(* IEC 61131-3 sources: daoli-st-library/DL_Motion (part 13) *)

(* ---- FB_DL_FilmWebCenter.st ---- *)
(*
    FB_DL_FilmWebCenter —— 膜卷纠偏（EPC）
    ------------------------------------------------------------------
    分类      : DL_Motion / Guide
    前缀      : FB_DL_
    版本      : 1.0.0
    溯源      : 纠偏为公开卷材处理工程结构（EPC / CPC：边缘或中心偏差 → 纠偏辊位置给定）；
                死区保持、断料保持、限速率、双侧行程钳位、错误分级与码位 100% 自有；
                与排线往复件、背隙修正件的职责严格分离（一个管横向对中、一个管往复排布、
                一个管传动链间隙）；clean-room 重写，未复制任何闭源厂商源码
    平台      : 纯 IEC 61131-3，CODESYS V3.5+ / TwinCAT 3 / InoProShop 通用
    作者      : 道莅代码库 · PLC编程专家（R19）
    ------------------------------------------------------------------
    功能说明  : 把边缘/中心偏差换算成纠偏辊位置给定。核心防御三条：
                ① 死区内保持——偏差在死区内给定不动，防辊子随噪声来回磨（不是把给定设成 0）；
                ② 限速率——纠偏动作过快会造成膜起皱甚至跑偏振荡；
                ③ 断料保持——膜断了还继续纠偏，辊子会一路顶到机械极限，复产后第一次穿膜
                   直接撞限位，故断料时给定保持末值、绝不追 0。
                其余防御：④ 行程域矛盾、增益或速率越域即故障级 02E4 并冻结在中心位
                   （增益过大是纠偏振荡的头号原因，硬限比「相信现场」更安全）；
                ⑤ 偏差非有限即故障级 02E5 并保持末次给定；
                ⑥ 给定双侧行程钳位，超限置 bLimited；⑦ 斜率限制首拍 fStep 由引脚换算，
                   不做除法；⑧ 状态机 CASE 含 ELSE 兜底，非法状态回 eIdle 并保持给定。
                职责边界：纠偏执行器的伺服闭环归驱动层，本件只出位置给定。
    错误码    : 16#0004_01D1 断料保持中 / 偏差在死区内给定保持——信息级，正常防御
                16#0004_01D2 预留禁用（信息级，不得挪用）
                16#0004_02E4 增益/速率/行程/采样参数非法——故障级，纠偏冻结在中心位
                16#0004_02E5 偏差输入非有限——故障级，给定保持末次有效
                16#0004_02E6 状态机落 ELSE 兜底（非法状态）——故障级，回 eIdle 并保持给定
    码位总账  : 16#0004_01D1 用 / 16#0004_01D2 预留 ｜ 16#0004_02E4 用 / 16#0004_02E5 用 / 16#0004_02E6 用
    状态机    : E_DL_WebState（eIdle / eManual / eAuto / eWebLost / eFault）五态，CASE 含 ELSE 兜底，
                ELSE 回 eIdle 并置故障级 02E6；失能不归零，只保持末值。
    采样约定  : fbTrigReset 在本体首部无条件刷新；速率步长由 tSampleTime 引脚换算；
                bInDeadband / bLimited / bWebLost 均为当拍组合量，不锁存。
    修订记录  : 2026-11-16 v1.0.0 首次入库（R19）
*)

(*
    枚举 : E_DL_WebState —— 纠偏工作状态（本文件为全库唯一属主）
*)
TYPE E_DL_WebState :
(
    eIdle    := 0,                            // 空闲：未使能，给定保持 / idle, disabled, the setpoint is held
    eManual  := 1,                            // 手动：走手动偏置给定 / manual, the setpoint follows the manual offset
    eAuto    := 2,                            // 自动：按偏差纠偏 / automatic, correcting by the measured deviation
    eWebLost := 3,                            // 断料：给定保持末值 / web lost, the setpoint holds its last value
    eFault   := 4                             // 故障：冻结在中心位 / fault, frozen at the centre
);
END_TYPE

FUNCTION_BLOCK FB_DL_FilmWebCenter
VAR_INPUT
    bEnable         : BOOL;                   // 使能，FALSE 输出保持末值（不归零）/ enable, FALSE holds the last setpoint without zeroing it
    bReset          : BOOL;                   // 复位，上升沿回中位并清状态 / reset, rising edge returns to the centre and clears the state
    bAuto           : BOOL := FALSE;          // TRUE = 自动纠偏，FALSE = 手动（走 fManualOffset）/ TRUE automatic, FALSE manual via the manual offset
    fDeviation      : REAL := 0.0;            // 边缘/中心偏差（正 = 偏向驱动侧）[mm] / edge or centre deviation, positive towards the drive side [mm]
    fGain           : REAL := 1.0;            // 偏差到位置给定增益 [mm/mm]，范围 0.1~20.0 / deviation to position gain [mm/mm], range 0.1~20.0
    fManualOffset   : REAL := 0.0;            // 手动偏置 [mm]，范围 fTravelMin~fTravelMax / manual offset [mm], range fTravelMin~fTravelMax
    fDeadband       : REAL := 0.3;            // 死区半宽 [mm]，范围 0.0~10.0 / deadband half width [mm], range 0.0~10.0
    fRateMax        : REAL := 5.0;            // 给定最大变化率 [mm/s]，范围 0.01~100.0 / maximum setpoint rate [mm/s], range 0.01~100.0
    fTravelMin      : REAL := -50.0;          // 行程下限 [mm] / travel lower bound [mm]
    fTravelMax      : REAL := 50.0;           // 行程上限 [mm]，必须 > fTravelMin / travel upper bound [mm], must be > fTravelMin
    bWebPresent     : BOOL := TRUE;           // 膜在位信号，FALSE = 断料 / web present signal, FALSE means the web is lost
    tSampleTime     : TIME := T#20MS;         // 采样周期 [ms]，范围 1~1000 / sample time [ms], range 1~1000
END_VAR
VAR_OUTPUT
    fPositionSp     : REAL;                   // 纠偏辊位置给定 [mm] / guide roller position setpoint [mm]
    bInDeadband     : BOOL;                   // 偏差在死区内（给定保持）/ the deviation is inside the deadband, the setpoint holds
    bLimited        : BOOL;                   // 受行程或速率限制 / limited by the travel or the rate
    bWebLost        : BOOL;                   // 断料保持中 / holding because the web is lost
    eErr            : UDINT;                  // 错误码，0=正常 / error id, 0=ok
    bError          : BOOL;                   // 故障标志，eErr 为故障级时 TRUE / error flag, TRUE on fault-level eErr
    bValid          : BOOL;                   // 给定是否可用 / setpoint valid flag
END_VAR
VAR
    fbTrigReset     : R_TRIG;                 // 复位上升沿实例，本体首部无条件刷新 / reset edge instance, refreshed unconditionally
    eState          : E_DL_WebState := eIdle; // 状态机当前态 / current state machine state
    fLastSp         : REAL;                   // 上一拍给定（斜率基准）[mm] / previous setpoint used by the ramp [mm]
    fTarget         : REAL;                   // 钳位与限速率前的目标给定 [mm] / target setpoint before clamping and ramping [mm]
    fStep           : REAL;                   // 本拍允许的最大变化量 [mm] / maximum allowed change in this cycle [mm]
    fDtSec          : REAL;                   // 采样周期秒值 [s] / sample time in seconds [s]
    fGainEff        : REAL;                   // 钳位后的增益 [mm/mm] / clamped gain [mm/mm]
    fDeadEff        : REAL;                   // 钳位后的死区半宽 [mm] / clamped deadband half width [mm]
    fManualEff      : REAL;                   // 钳位后的手动偏置 [mm] / clamped manual offset [mm]
    nDtMs           : DINT;                   // 采样周期毫秒整数 [ms] / sample time in integer milliseconds [ms]
    bInit           : BOOL := FALSE;          // 首扫标志，初值 FALSE，判据 NOT bInit / first-scan flag, initial FALSE, tested with NOT
END_VAR
VAR CONSTANT
    DL_EPC_GAIN_MIN  : REAL := 0.1;           // 增益下限 [mm/mm] / gain lower bound [mm/mm]
    DL_EPC_GAIN_MAX  : REAL := 20.0;          // 增益上限 [mm/mm] / gain upper bound [mm/mm]
    DL_EPC_RATE_MIN  : REAL := 0.01;          // 速率下限 [mm/s] / rate lower bound [mm/s]
    DL_EPC_RATE_MAX  : REAL := 100.0;         // 速率上限 [mm/s] / rate upper bound [mm/s]
    DL_EPC_DB_MAX    : REAL := 10.0;          // 死区半宽上限 [mm] / deadband half width upper bound [mm]
    DL_EPC_DT_MAX    : TIME := T#1S;          // 采样周期上限 [ms] / sample time upper bound [ms]
    DL_EPC_DT_MIN    : TIME := T#1MS;         // 采样周期下限 [ms] / sample time lower bound [ms]
    DL_FLOAT_EPS     : REAL := 1.0E-6;        // 浮点判等容差 [无量纲] / float equality tolerance [dimensionless]
    DL_EPC_MS_PER_S  : REAL := 1000.0;        // 毫秒到秒换算因子 [ms/s] / milliseconds per second [ms/s]
    DL_EPC_INF_GUARD : REAL := 1.0E38;        // 非有限幅值判定阈值 [无量纲] / non-finite magnitude guard [dimensionless]
    DL_EPC_ZERO      : REAL := 0.0;           // 零值常量，避免裸字面量 [mm] / zero constant, avoids a bare literal [mm]
END_VAR

// 段 1｜边沿实例无条件周期刷新（红线：严禁放入条件分支）/ segment 1, unconditional edge refresh
fbTrigReset(CLK := bReset);

// 段 2｜输出与错误状态预置（fPositionSp 为保持量，故障与断料时均保持）/ segment 2, preset outputs, the setpoint is held
eErr := 0;                                    // 预置无错误 / preset no error
bError := FALSE;                              // 预置无故障 / preset no fault
bInDeadband := FALSE;                         // 预置非死区 / preset outside the deadband
bLimited := FALSE;                            // 预置未受限 / preset not limited
bWebLost := NOT bWebPresent;                  // 断料标志由在位信号导出 / the web lost flag derives from the present signal

// 段 3｜首扫初始化（唯一合法范式：初值 FALSE，判据 NOT bInit）/ segment 3, first-scan initialisation
IF NOT bInit THEN
    fLastSp := DL_EPC_ZERO;                   // 首扫给定基准取中心位 / the setpoint reference starts at the centre
    bInit := TRUE;                            // 首扫只做一次 / first scan runs once only
END_IF

// 段 4｜参数闸：行程域、增益、速率、采样周期（任一非法即冻结在中心位）/ segment 4, parameter gate
IF (fTravelMax <= fTravelMin)
   OR (fGain < DL_EPC_GAIN_MIN) OR (fGain > DL_EPC_GAIN_MAX)
   OR (fRateMax < DL_EPC_RATE_MIN) OR (fRateMax > DL_EPC_RATE_MAX)
   OR (tSampleTime < DL_EPC_DT_MIN) OR (tSampleTime > DL_EPC_DT_MAX) THEN
    eErr := 16#0004_02E4;                     // 参数非法故障码 / illegal parameter fault id
    bError := TRUE;                           // 置故障标志 / raise the error flag
    eState := eFault;                         // 落故障态 / enter the fault state
    fPositionSp := DL_EPC_ZERO;               // 冻结在中心位（唯一安全的固定点）/ freeze at the centre, the only safe fixed point
    bValid := FALSE;                          // 给定不可用 / the setpoint is not usable
    RETURN;                                   // 故障级提前返回 / early return on fault
END_IF

// 段 5｜偏差非有限闸：给定保持末次有效（绝不追 0）/ segment 5, non-finite gate holds the setpoint
IF (fDeviation <> fDeviation) OR (fDeviation > DL_EPC_INF_GUARD) OR (fDeviation < -DL_EPC_INF_GUARD) THEN
    eErr := 16#0004_02E5;                     // 偏差非有限故障码 / non-finite deviation fault id
    bError := TRUE;                           // 置故障标志 / raise the error flag
    eState := eFault;                         // 落故障态 / enter the fault state
    fPositionSp := fLastSp;                   // 保持末次给定 / hold the last setpoint
    bValid := FALSE;                          // 给定不可用 / the setpoint is not usable
    RETURN;                                   // 故障级提前返回 / early return on fault
END_IF

// 段 6｜域钳位与速率步长（无历史依赖，不做除法）/ segment 6, domain clamp and rate step
fGainEff := fGain;                            // 增益已由段 4 保证在域内 / the gain is already in range by segment 4
fDeadEff := MIN(MAX(fDeadband, DL_EPC_ZERO), DL_EPC_DB_MAX); // 死区半宽收敛到 0.0~10.0 mm / converge the deadband into 0.0~10.0 mm
fManualEff := MIN(MAX(fManualOffset, fTravelMin), fTravelMax); // 手动偏置收敛到行程域 / converge the manual offset into the travel range
nDtMs := TIME_TO_DINT(tSampleTime);           // 采样周期整数毫秒 [ms] / sample time in integer milliseconds [ms]
fDtSec := DINT_TO_REAL(nDtMs) / DL_EPC_MS_PER_S; // 换算为秒，除子为常量 [s] / convert to seconds, the divisor is a constant [s]
fStep := fRateMax * fDtSec;                   // 本拍允许的最大变化量 [mm] / maximum allowed change in this cycle [mm]

// 段 7｜复位沿：回中位并清状态 / segment 7, reset returns to the centre
IF fbTrigReset.Q THEN
    fLastSp := DL_EPC_ZERO;                   // 给定基准回中心位 / the setpoint reference returns to the centre
    fPositionSp := DL_EPC_ZERO;               // 给定回中位 / the setpoint returns to the centre
    IF eState = eFault THEN
        eState := eIdle;                      // 故障态允许由复位退出 / a reset leaves the fault state
    END_IF
END_IF

// 段 8｜状态选择（断料优先级最高，其次使能与手自动）/ segment 8, state selection
IF NOT bWebPresent THEN
    eState := eWebLost;                       // 断料优先，给定保持 / web loss has the highest priority, the setpoint holds
    bWebLost := TRUE;                         // 发布断料标志 / publish the web lost flag
ELSE
    bWebLost := FALSE;                        // 在位则清断料标志 / clear the flag when the web is present
    IF eState = eWebLost THEN
        eState := eIdle;                      // 断料解除回空闲，由使能重新决定手自动 / leaving the web lost state returns to idle
    END_IF
END_IF
IF (eState <> eWebLost) AND (eState <> eFault) THEN
    IF NOT bEnable THEN
        eState := eIdle;                      // 失能回空闲（保持不归零）/ disabled returns to idle without zeroing the setpoint
    ELSIF bAuto THEN
        eState := eAuto;                      // 自动纠偏 / automatic correction
    ELSE
        eState := eManual;                    // 手动偏置 / manual offset
    END_IF
END_IF

// 段 9｜目标给定（含死区保持与断料保持）/ segment 9, target setpoint with deadband and web loss holding
CASE eState OF
    eIdle:
        fTarget := fLastSp;                   // 空闲保持末值，不归零 / idle holds the last value without zeroing it

    eManual:
        fTarget := fManualEff;                // 手动走偏置给定 / manual follows the offset

    eAuto:
        IF ABS(fDeviation) <= fDeadEff THEN
            fTarget := fLastSp;               // 死区内保持，绝不设成 0 / hold inside the deadband, never set it to zero
            bInDeadband := TRUE;              // 发布死区标志 / publish the deadband flag
            eErr := 16#0004_01D1;             // 信息级：偏差在死区内给定保持 / info level, the setpoint holds inside the deadband
        ELSE
            fTarget := fLastSp + fGainEff * fDeviation; // 增量式纠偏：在上一拍给定上叠加 / incremental correction on top of the previous setpoint
        END_IF

    eWebLost:
        fTarget := fLastSp;                   // 断料保持末值 / web lost holds the last value
        eErr := 16#0004_01D1;                 // 信息级：断料保持中 / info level, holding because the web is lost

    eFault:
        fTarget := fLastSp;                   // 故障态保持末值 / the fault state holds the last value

ELSE
    eErr := 16#0004_02E6;                     // 故障级：非法状态兜底 / fault level, illegal state fallback
    bError := TRUE;                           // 置故障标志 / raise the error flag
    eState := eIdle;                          // 回空闲态 / fall back to idle
    fTarget := fLastSp;                       // 保持末值，不产生跳变 / hold the last value, no jump
END_CASE

// 段 10｜行程双侧钳位（只做单侧是常见缺陷）/ segment 10, two-sided travel clamp
IF fTarget > fTravelMax THEN
    fTarget := fTravelMax;                    // 上限钳位 / clamp at the upper bound
    bLimited := TRUE;                         // 标记行程受限 / flag the travel limit
ELSIF fTarget < fTravelMin THEN
    fTarget := fTravelMin;                    // 下限钳位 / clamp at the lower bound
    bLimited := TRUE;                         // 标记行程受限 / flag the travel limit
END_IF

// 段 11｜限速率（每拍最多变化 fStep，防膜起皱与跑偏振荡）/ segment 11, rate limiting
IF fStep > DL_EPC_ZERO THEN
    IF fTarget > (fLastSp + fStep) THEN
        fTarget := fLastSp + fStep;           // 正向每拍限幅 / limit the positive step per cycle
        bLimited := TRUE;                     // 标记速率受限 / flag the rate limit
    ELSIF fTarget < (fLastSp - fStep) THEN
        fTarget := fLastSp - fStep;           // 负向每拍限幅 / limit the negative step per cycle
        bLimited := TRUE;                     // 标记速率受限 / flag the rate limit
    END_IF
END_IF

// 段 12｜发布给定 / segment 12, publish the setpoint
fPositionSp := fTarget;                       // 输出纠偏辊位置给定 [mm] / publish the guide roller setpoint [mm]
fLastSp := fTarget;                           // 记录为下一拍斜率基准 / remember it as the next ramp reference
IF NOT bError THEN
    bValid := TRUE;                           // 无故障则给定可用 / usable when no fault is present
END_IF
END_FUNCTION_BLOCK

(* ---- FB_DL_FlyingCutSync.st ---- *)
(*
  FB_DL_FlyingCutSync  —  飞剪同步切（相位取模 / 切窗判据 / 电子齿轮追赶 / 单拍下刀）/ Flying-cut synchronisation
  分类 Category : DL_Motion
  码位 Code     : 16#04_0_A3
  版本 Version  : 1.0.1
  来源 Source   : t1-6-plcopen — IEC 61131-3 标准语义的道莅防御性实现
  溯源 Origin   : PLCopen 飞剪/电子齿轮公开语义借鉴，clean-room 实现，仅借相位取模与切窗概念，未复制源码行
  功能 Function : 1) 主轴位置对 fCutLengthMm 取模（FLOOR 口径，负向同样收敛）得切长相位 fPhaseMm；
                  2) 相位落在 [fSyncWindowStartMm, fSyncWindowEndMm] 内置 bInSyncWindow，窗口内方允许下刀；
                  3) 同步误差 fSyncErrorMm = 刀轴位置 − 相位 × fCutOverlapRatio，进 fSyncTolMm 才发下刀脉冲；
                  4) 下刀脉冲 bCutCmd 为**单拍脉冲**（脉冲语义：置位 1 个 PLC 周期），由内部 _bCutPulse 置位、
                     段 8 统一出口映射，次拍段 1 清零，绝不在 CASE 内二次写输出（N2 / R187①）；
                  5) 切完按 tCutDwell 保压（刀在料内停留），保压结束进回程相，等相位越过窗尾再回等待相；
                  6) 每圈只允许一刀：以圈索引 fTurnsInt 与 _nCutTurnIdx 比较做单圈互锁（防同圈重刀）。
  边界 Boundary : ① fCutLengthMm <= 0 判组态错（取模除零前置，R45）；窗口起止倒置或宽 <= 0 判组态错且不运行；
                      fSyncTolMm <= 0 / fCutOverlapRatio <= 0 同判组态错，码 00A3，状态进 eFault；
                  ② 未同步时**禁止** bCutCmd：互锁写在件内（窗口 + 容差 + 单圈 + 主轴正向四条件同时成立），
                     不外抛给上层组合逻辑（防上层漏联锁切刀撞料）；
                  ③ nCutCount 到 uCountPreset 后 bPresetReached 置位；计数在 UDINT 上限前饱和**不回绕**，
                     预置比较用「增量前预判」而非事后比较（不给 TRUNC(x)+1 型写法，R28-3）；
                  ④ 切窗内主轴反转立即判废并置 01A3（反转期刀轴与料带速度矢量相反，下刀即撕料）；
                  ⑤ uCountPreset = 0 视为「不启用预置」：bPresetReached 恒 FALSE，置信息级 07A3；
                  ⑥ 解除路径自证：_bFault 清除 = rtReset.Q（引脚可满足）；01A3 另可由「主轴恢复正向
                     且相位出新窗」按码专清（两路径互不掩盖，R188）。
  依赖 Depends  : I_DL_MotionAxis / E_DL_AxisState（DL_Motion 既有契约件，零修改，只注入不实例化）；
                  仅 Standard.library（TON / R_TRIG / ABS / MIN / MAX）
  同拍双窗配比  : tCutDwell（刀内停留）与 tonGuard 自复位心跳窗不同源；配比约束
                  tCutDwell <= DL_GUARD_WINDOW / 2，保证保压段内至少一次心跳判活（R100）

  码表 Error codes（本件格 04_0_A3，子码步进 +0x10）:
    16#0004_00A3 故障级：组态非法（切长 <= 0 / 窗口倒置或宽 <= 0 / 容差 <= 0 / 重叠比 <= 0）
    16#0004_01A3 故障级：切窗内主轴反转，本次切割判废
    16#0004_03A3 故障级：状态机落 ELSE 兜底（非法相位 ID）
    16#0004_04A3 信息级：下刀脉冲已发出（bCutCmd 单拍同源，不置 bError）
    16#0004_05A3 信息级：切割计数达预置（bPresetReached 同拍置位，不置 bError）
    16#0004_06A3 信息级：切窗内同步超差，本次跳过不下刀（互锁生效，不置 bError）
    16#0004_07A3 信息级：预置计数未组态（uCountPreset = 0，预置出口恒 FALSE）

  修订历史 Revision :
    2026-11-18  v1.0.0  R37 首版
*)

TYPE E_DL_FlyingCutState :
(
    eIdle       := 0,   // 空闲：未使能，不出切窗判据 / Idle, no window evaluation while disabled
    eWaiting    := 10,  // 等待：等相位进入切窗 / Waiting for the phase to enter the cut window
    eSyncWindow := 20,  // 窗内：按容差追赶，达标即下刀 / Inside the window, chasing the tolerance
    eCutting    := 30,  // 切割：刀在料内保压（tCutDwell）/ Cutting, the knife dwells inside the web
    eReturning  := 40,  // 回程：等相位越过窗尾，准备下一圈 / Returning, waiting for the phase to pass the window end
    eFault      := 90   // 故障：组态非法或反转判废锁定 / Fault, illegal configuration or a latched reversal reject
);
END_TYPE

FUNCTION_BLOCK FB_DL_FlyingCutSync
VAR_INPUT
    bEnable        : BOOL := FALSE;              // 总使能，FALSE 时禁止下刀 / Master enable, a low level forbids cutting
    bReset         : BOOL := FALSE;              // 复位，上升沿清故障锁存 / Reset, rising edge clears the latch
    fCutLengthMm   : REAL := 1000.0;             // 单刀切长（取模基数）[mm]，域 > 0 / Cut length, the modulo base [mm]
    fSyncWindowStartMm : REAL := 5.0;            // 切窗起点相位 [mm]，域 >= 0 / Window start phase [mm]
    fSyncWindowEndMm   : REAL := 45.0;           // 切窗终点相位 [mm]，须 > 起点 / Window end phase [mm]
    fCutOverlapRatio   : REAL := 1.0;            // 刀轴等效行程与相位之比 [1]，域 > 0 / Knife travel per phase unit [1]
    tCutDwell      : TIME := T#120MS;            // 刀内保压时间 [ms]，域 > 0 / Knife dwell inside the web [ms]
    fSyncTolMm     : REAL := 0.5;                // 允许下刀的同步误差 [mm]，域 > 0 / Sync tolerance permitting a cut [mm]
    uCountPreset   : UDINT := 10000;             // 切割计数预置 [次]，0 = 不启用预置 / Cut count preset, zero disables it
END_VAR
VAR_OUTPUT
    bCutCmd        : BOOL;                       // 下刀指令（脉冲语义：置位 1 个 PLC 周期）/ Cut command, asserted for exactly one PLC scan
    bInSyncWindow  : BOOL;                       // 相位处于切窗内 / Phase inside the cut window
    fSyncErrorMm   : REAL;                       // 同步误差 [mm]，刀轴位置 − 相位×重叠比 / Sync error [mm]
    fPhaseMm       : REAL;                       // 当前切长相位 [mm]，域 [0, fCutLengthMm) / Present phase inside one cut [mm]
    nCutCount      : UDINT;                      // 累计切割次数 [次]，饱和不回绕 / Accumulated cut count, saturated, never wrapped
    bPresetReached : BOOL;                       // 计数达预置标志（保持型）/ Preset reached flag, held
    bValid         : BOOL;                       // 判据可用标志 / Criteria usable
    bError         : BOOL;                       // 故障标志，派生自锁存 / Fault flag derived from the latch
    nErrId         : UDINT;                      // 事件码，0 = 无事件 / Event code, 0 = no event
    eStateOut      : E_DL_FlyingCutState;        // 状态出口，段尾单点映射 / State outlet, mapped at the tail
END_VAR
VAR_IN_OUT
    iMasterAxis    : I_DL_MotionAxis;            // 料带线轴接口引用（注入，不实例化）/ Web master axis reference, injected
    iCutAxis       : I_DL_MotionAxis;            // 刀轴接口引用（注入，不实例化）/ Knife axis reference, injected
END_VAR
VAR
    tonDwell       : TON;                        // 刀内保压计时，每拍无条件调用 / Knife dwell timer, called unconditionally
    tonGuard       : TON;                        // 周期心跳窗，自复位 / Periodic guard window, self-resetting
    rtReset        : R_TRIG;                     // 复位上升沿 / Reset rising edge
    _eState        : E_DL_FlyingCutState := E_DL_FlyingCutState.eIdle;  // 内部相位（CASE 唯一写入目标）/ Internal phase
    _uFault        : UDINT;                      // 故障码锁存 / Latched fault code
    _uInfo         : UDINT;                      // 信息码，每拍重算 / Information code, recomputed per scan
    _bFault        : BOOL;                       // 故障锁存位 / Latched fault bit
    _bParamBad     : BOOL;                       // 组态非法聚合 / Configuration invalid aggregate
    _bCutPulse     : BOOL;                       // 内部下刀单拍标志 → 段 8 映射 / Internal one-shot cut flag
    _bPresetReached: BOOL;                       // 预置到达保持量 / Held preset-reached value
    _bSameTurn     : BOOL;                       // 本圈已下刀（单圈互锁）/ A cut already happened in this turn
    _bWindowNow    : BOOL;                       // 本拍窗内判据 / Window predicate this scan
    _bReverse      : BOOL;                       // 切窗内主轴反转 / Master reversal inside the window
    _fTurns        : REAL;                       // 位置除切长的商（圈数，实数）/ Turn count as a real quotient
    _fPhase        : REAL;                       // 切长相位 [mm] / Phase inside one cut [mm]
    _fSyncErr      : REAL;                       // 同步误差 [mm] / Sync error [mm]
    _fExpPos       : REAL;                       // 刀轴期望等效行程 [mm] / Expected knife equivalent travel [mm]
    _dTurnsInt     : DINT;                       // FLOOR 后的圈索引（负向同样收敛）/ Floor turn index, negative safe
    _uCountAcc     : UDINT;                      // 计数保持量 [次] / Held count value
    _nCutTurnIdx   : DINT := -1;                 // 最后一次下刀的圈索引（-1=尚无下刀，防初值吃首圈）/ Turn index, -1 = none yet
    _bGuardBreak   : BOOL := TRUE;               // 心跳窗断输入一拍 / One-scan guard break
END_VAR
VAR CONSTANT
    DL_CNT_MAX     : UDINT := 16#FFFF_FFFE;      // 计数饱和上限（留 1 位防溢出）[次] / Saturation ceiling, one below the wrap
    DL_EPS         : REAL  := 1.0E-6;            // 判零容差 [1] / Zero tolerance
    DL_GUARD_WINDOW : TIME := T#2S;              // 心跳观察窗 [ms]，自复位节拍 / Guard window, self-resetting
    DL_WIN_MAX_MM  : REAL  := 1.0E6;             // 相位与搜索量绝对值上限 [mm] / Magnitude ceiling for phases [mm]
END_VAR

(* —— 段 0：定时器与边缘检测无条件周期刷新（R182：调用语句本身不得置于 IF 内） —— *)
rtReset(CLK := bReset);                                          // 复位上升沿，每拍必调
tonGuard(IN := (NOT tonGuard.Q) AND (NOT _bGuardBreak), PT := DL_GUARD_WINDOW);  // 心跳窗自复位
_bGuardBreak := FALSE;                                           // 断输入拍在调用后自清
tonDwell(IN := (_eState = E_DL_FlyingCutState.eCutting), PT := tCutDwell);       // 保压计时（表达式入参）

(* —— 段 1：单拍量预清零（计数 / 预置 / 锁存不入清单，R187①） —— *)
_uInfo   := 16#0000_0000;   // 信息码每拍重算
bError   := FALSE;          // 故障出口每拍重算，段 7 由锁存派生
bValid   := FALSE;          // 判据可用缺省 FALSE
bCutCmd  := FALSE;          // 下刀出口缺省 FALSE（段 8 单点映射，脉冲宽度 = 1 拍）
_bCutPulse := FALSE;        // 内部下刀单拍标志预清零
_bParamBad := FALSE;        // 组态非法预清零
_bWindowNow := FALSE;       // 窗内判据预清零
_bReverse := FALSE;         // 反转标志预清零
_bSameTurn := FALSE;        // 单圈互锁标志预清零

(* —— 段 2：复位沿清锁存（按码专清 + 恢复沿清码，R188） —— *)
IF rtReset.Q THEN
    _bFault := FALSE;            // 复位沿清锁存位
    _uFault := 16#0000_0000;     // 复位沿清锁存码
END_IF

(* —— 段 3：组态域闸（覆盖全部参与判据换算的引脚，R151） —— *)
IF (fCutLengthMm <> fCutLengthMm) OR (fCutLengthMm <= 0.0) OR (fCutLengthMm > DL_WIN_MAX_MM) THEN
    _bParamBad := TRUE;          // 切长非法：取模除零前置（R45）
END_IF
IF (fSyncWindowStartMm <> fSyncWindowStartMm) OR (fSyncWindowStartMm < 0.0) THEN
    _bParamBad := TRUE;          // 窗起点非法
END_IF
IF (fSyncWindowEndMm <> fSyncWindowEndMm) OR (fSyncWindowEndMm <= fSyncWindowStartMm) THEN
    _bParamBad := TRUE;          // 窗止倒置或宽度 <= 0
END_IF
IF (NOT _bParamBad) AND ((fSyncWindowEndMm - fSyncWindowStartMm) <= 0.0) THEN
    _bParamBad := TRUE;          // 窗宽 <= 0（显式复检，防浮点相消导致宽度判据静默失效）
END_IF
IF (fSyncTolMm <> fSyncTolMm) OR (fSyncTolMm <= 0.0) THEN
    _bParamBad := TRUE;          // 同步容差非法（互锁门限为 0 等于永不下刀）
END_IF
IF (fCutOverlapRatio <> fCutOverlapRatio) OR (fCutOverlapRatio <= 0.0) THEN
    _bParamBad := TRUE;          // 重叠比非法（期望行程的比例因子）
END_IF
IF TIME_TO_DINT(tCutDwell) <= 0 THEN
    _bParamBad := TRUE;          // 保压时间非法（零保压会让刀在料内瞬时撤回）
END_IF
IF _bParamBad THEN
    _uFault := 16#0004_00A3;     // 故障级：组态非法
    _bFault := TRUE;             // 锁存位置位（复位沿可清）
    bError  := TRUE;             // 故障标志置位（R45 配对）
    _eState := E_DL_FlyingCutState.eFault;  // 状态机进故障相
END_IF

(* —— 段 4：相位取模与同步误差（仅无组态错时计算） —— *)
IF NOT _bParamBad THEN
    _fTurns := iMasterAxis.fPosition / fCutLengthMm;               // 圈数商（分母已证 > 0）
    _dTurnsInt := REAL_TO_DINT(_fTurns);                           // 向零截断
    IF (_fTurns < 0.0) AND (ABS(_fTurns - DINT_TO_REAL(_dTurnsInt)) > DL_EPS) THEN
        _dTurnsInt := _dTurnsInt - 1;                              // 负向修正为 FLOOR，保证相位恒 >= 0
    END_IF
    _fPhase := iMasterAxis.fPosition - (DINT_TO_REAL(_dTurnsInt) * fCutLengthMm);  // 切长相位 [mm]
    IF _fPhase < 0.0 THEN
        _fPhase := _fPhase + fCutLengthMm;                         // 相消残差归正（浮点尾差兜底）
    END_IF
    IF _fPhase >= fCutLengthMm THEN
        _fPhase := _fPhase - fCutLengthMm;                         // 上行越界折回一格
    END_IF
    _bWindowNow := (_fPhase >= fSyncWindowStartMm) AND (_fPhase <= fSyncWindowEndMm);  // 窗内判据
    _fExpPos := _fPhase * fCutOverlapRatio;                        // 刀轴期望等效行程 [mm]
    _fSyncErr := iCutAxis.fPosition - _fExpPos;                    // 同步误差 [mm]
    IF _bWindowNow AND (iMasterAxis.fVelocity < -DL_EPS) THEN
        _bReverse := TRUE;                                         // 窗内主轴反转：判废
    END_IF
    IF _dTurnsInt = _nCutTurnIdx THEN
        _bSameTurn := TRUE;                                        // 本圈已下刀：单圈互锁生效
    END_IF
    fPhaseMm     := _fPhase;                                       // 相位出口
    fSyncErrorMm := _fSyncErr;                                     // 误差出口
END_IF
bInSyncWindow := _bWindowNow;                                      // 窗内出口（诊断与上层互锁共用）

(* 段 4B｜按码专清：01A3 的恢复沿条件依赖本拍相位与速度，故必须置于段 4 之后判（R188 可达清除边） *)
IF (_uFault = 16#0004_01A3) AND _bFault AND (iMasterAxis.fVelocity > DL_EPS) AND (NOT _bWindowNow) THEN
    _uFault := 16#0000_0000;          // 主轴恢复正向且相位已出新窗：反转判废可解
    _bFault := FALSE;                 // 锁存位同步清（与 rtReset.Q 路径互不掩盖）
END_IF

(* —— 段 5：相位机（只做迁移与内部单拍标志；输出在段 8） —— *)
CASE _eState OF

E_DL_FlyingCutState.eIdle:
    IF bEnable AND (NOT _bFault) AND (NOT _bParamBad) THEN
        _eState := E_DL_FlyingCutState.eWaiting;                   // 使能且无故障：进等待相
    END_IF

E_DL_FlyingCutState.eWaiting:
    IF (NOT bEnable) THEN
        _eState := E_DL_FlyingCutState.eIdle;                      // 失能：回空闲，禁止下刀
    ELSIF _bReverse THEN
        _uFault := 16#0004_01A3;                                   // 故障级：切窗内主轴反转
        _bFault := TRUE;                                           // 锁存
        bError  := TRUE;                                           // 故障标志置位（R45 配对）
        _eState := E_DL_FlyingCutState.eFault;                     // 进故障相
    ELSIF _bWindowNow THEN
        _eState := E_DL_FlyingCutState.eSyncWindow;                // 进窗：开始追赶
    END_IF

E_DL_FlyingCutState.eSyncWindow:
    IF (NOT bEnable) THEN
        _eState := E_DL_FlyingCutState.eIdle;                      // 失能：退出窗内（不下刀）
    ELSIF _bReverse THEN
        _uFault := 16#0004_01A3;                                   // 故障级：切窗内主轴反转
        _bFault := TRUE;                                           // 锁存
        bError  := TRUE;                                           // 故障标志置位（R45 配对）
        _eState := E_DL_FlyingCutState.eFault;                     // 进故障相
    ELSIF NOT _bWindowNow THEN
        _uInfo := 16#0004_06A3;                                    // 信息级：出窗未达容差，本次跳过
        _eState := E_DL_FlyingCutState.eWaiting;                    // 回等待相，等下一圈
    ELSIF _bSameTurn THEN
        _eState := E_DL_FlyingCutState.eWaiting;                    // 本圈已切：不许重刀，回等待
    ELSIF ABS(_fSyncErr) <= fSyncTolMm THEN
        _bCutPulse := TRUE;                                        // 四条件同时成立：置内部下刀单拍
        _nCutTurnIdx := _dTurnsInt;                                // 记录本圈已下刀（单圈互锁）
        _eState := E_DL_FlyingCutState.eCutting;                   // 进保压相
        _bGuardBreak := TRUE;                                      // 心跳窗重启（保压段重新判活）
        IF _uCountAcc < DL_CNT_MAX THEN
            _uCountAcc := _uCountAcc + 1;                          // 计数 +1（饱和不回绕，R28-3）
        END_IF
        IF (uCountPreset > 0) AND (_uCountAcc >= uCountPreset) THEN
            IF NOT _bPresetReached THEN
                _uInfo := 16#0004_05A3;                            // 信息级：计数达预置（首次置位拍）
            END_IF
            _bPresetReached := TRUE;                               // 预置到达保持量置位
        END_IF
    ELSE
        _uInfo := 16#0004_06A3;                                    // 信息级：窗内同步超差，互锁生效不下刀
    END_IF

E_DL_FlyingCutState.eCutting:
    IF tonDwell.Q THEN
        _eState := E_DL_FlyingCutState.eReturning;                 // 保压完成：进回程相
    END_IF

E_DL_FlyingCutState.eReturning:
    IF (NOT bEnable) THEN
        _eState := E_DL_FlyingCutState.eIdle;                      // 失能：回空闲
    ELSIF (_fPhase > fSyncWindowEndMm) OR (_fPhase < fSyncWindowStartMm) THEN
        _eState := E_DL_FlyingCutState.eWaiting;                   // 相位已出窗：回等待相等下一圈
    END_IF

E_DL_FlyingCutState.eFault:
    IF (NOT _bFault) AND (NOT _bParamBad) AND bEnable THEN
        _eState := E_DL_FlyingCutState.eWaiting;                   // 锁存已清且组态合法：回等待相
    END_IF

ELSE
    _uFault := 16#0004_03A3;                                       // 故障级：相位 ID 越界（枚举兜底）
    _bFault := TRUE;                                               // 锁存
    bError  := TRUE;                                               // 故障标志置位（R45 配对）
    _eState := E_DL_FlyingCutState.eFault;                         // 强制回故障相
END_CASE

(* —— 段 6：预置比较（保持量推进 + 计数上限兜底，禁 TRUNC(x)+1 型写法） —— *)
IF uCountPreset = 0 THEN
    _bPresetReached := FALSE;             // 未组态预置：出口恒 FALSE（不做数值比较）
    _uInfo := 16#0004_07A3;               // 信息级：预置未组态
ELSIF _uCountAcc >= uCountPreset THEN
    _bPresetReached := TRUE;              // 已达预置：保持置位（不随计数变化回落）
END_IF

(* —— 段 7：故障码优先级链（每个 bError 置位源在此均有码，R45 配对） —— *)
IF _bParamBad THEN
    _uFault := 16#0004_00A3;              // 组态非法优先上报（其余码不得掩盖）
    _bFault := TRUE;                      // 锁存
    bError  := TRUE;                      // 故障标志置位
END_IF

(* —— 段 8：出口单点映射（名实同源；脉冲两段式已在段 1 与段 5 完成） —— *)
bCutCmd        := _bCutPulse;             // 下刀出口：仅本拍置位，宽度恰 1 个 PLC 周期
nCutCount      := _uCountAcc;             // 计数出口
bPresetReached := _bPresetReached;        // 预置出口（保持型）
eStateOut      := _eState;                // 状态出口
IF _bFault THEN
    nErrId := _uFault;                    // 故障锁存码回放（不在故障相按当下输入重推）
    bError := TRUE;                       // 故障出口派生自锁存
ELSE
    nErrId := _uInfo;                     // 信息码
END_IF
bValid := bEnable AND (NOT _bFault) AND (NOT _bParamBad);  // 判据可用：使能且无故障且组态合法

END_FUNCTION_BLOCK

(* ---- FB_DL_FlyingSawSyncSeq.st ---- *)
//==============================================================================
// 功能块：FB_DL_FlyingSawSyncSeq ｜ 中文名称：飞锯同步切入-切割-返回全序列
// 所属子库：DL_Motion ｜ 版本：v1.0.1 ｜ 日期：2026-11-23
// 兼容：CODESYS V3.5+ / TwinCAT 3 / 汇川 InoProShop（纯 IEC 61131-3 第 3 版，零方言）
// 功能描述：飞锯电子凸轮全序列编排。以同步轴（主轴）位置为时间基准：在切割
//           锚点前方 fSyncLen 区间内把主从速比从 0 线性爬升到 1（同步切入），
//           保持速比 1 走完 fCutLen 切割窗口（本窗内 bCutReq 置位），再对称
//           降回 0（同步返回）。速比全部按主轴位置增量生成，即相对同步轴
//           补偿：主轴中途变速不破坏同步关系，刀轴速度 = 主轴速度 × fRatio。
// 开源溯源 (Origin)：原创实现（t1-6-plcopen 运动序列语义深化 + S-9 工程惯例，
//           零外部源码行，clean-room 独立编写）
// 公开接口清单：输入 bEn / bStart / fMasterPos / fSyncLen / fCutLen；
//               输出 bKnifeRun / fRatio / bCutReq / bCycleDone / eState /
//               uErrCode / bValid
// 单位表：fMasterPos[mm] / fSyncLen[mm] / fCutLen[mm] / fRatio[1]（无量纲比）
// 输入契约：fMasterPos 为主轴编码器工程位置，须单调正向为切割方向；fSyncLen
//           /fCutLen 为工艺给定窗长，启动闸拒绝非正值；bStart 沿触发单周期。
// 输出契约：fRatio 注入刀轴速度合成（刀速 = 主速 × fRatio）；bCutReq 为
//           请求级信号（非执行器驱动级）；bCycleDone 单拍计件脉冲；
//           uErrCode 信息级不锁存；bValid = FALSE 拍全部输出视为不可信。
// 错误码表：16#0004_08C0 信息级（参数非法拒绝启动、输入非有限安全侧回怠速、
//           序列中途参数退化中止，不置 bError）/
//           16#0004_08C1 预留禁用（不得挪用）
// 状态机：E_DL_FlyingSawState（本文件唯一定义，全库唯一属主）：
//           eIdle = 0 / eWait = 10 / eSyncIn = 20 / eCutting = 30 / eSyncOut = 40
// 边界行为：① fSyncLen / fCutLen <= 0 或非有限 → 拒绝启动（怠速态）+ 信息码；
//           ② 主轴位置非有限 → 速比冻结 0、序列中止回 eIdle（安全侧）；
//           ③ 速比全程钳 0..1，除法分母 fSyncLen 先过正域闸；
//           ④ 切入相内主轴位置跳变已越锚点 → 相位判据顺带直入切割相不丢拍
//             （未来窗锚点下，启动沿不可能已越窗）；
//           ⑤ CASE 带 ELSE 非法状态兜底回 eIdle；
//           ⑥ R_TRIG 每拍无条件刷新（不入分支，红线 R7）；
//           ⑦ bCycleDone 两段式单拍脉冲（内部置位 → 统一出口映射）；
//           ⑧ 活动相内主轴位置倒退超容差（方向反转）→ 序列中止回怠速，
//             信息级 08C0 复用留痕（R90），速比归零安全侧。
// 修订历史：v1.0.0 2026-11-23 首版（R73 派单 · 批 1 · 序 1）
//           v1.0.1 2026-11-23 R73 返修：锚点改未来窗语义——启动沿锁存
//           fAnchor := fMasterPos + fSyncLen（预留一个同步窗长的提前量），
//           切入窗 [fAnchor−fSyncLen, fAnchor] 整体落在主轴前方，速比
//           0→1 爬坡真实发生；bCutReq 仍仅在速比 1 切割相内置位（头注释
//           与实现保持一致，R372 语料保真）。
//==============================================================================

(*------------------------------------------------------------------------------
 * 枚举: E_DL_FlyingSawState（归属本功能块，同文件发布，全库唯一属主）
 * 含义: 飞锯序列相位，成员与 CASE 标签双向完备。
 *-----------------------------------------------------------------------------*)
TYPE E_DL_FlyingSawState :
(
    eIdle    := 0,    // 怠速：速比 0，等待启动沿 / Idle, ratio 0, waiting for start edge
    eWait    := 10,   // 待同步：锚点已记，等主轴进入同步窗 / Waiting, anchor set, master not yet in sync window
    eSyncIn  := 20,   // 同步切入：速比 0→1 线性爬升 / Sync-in, ratio ramping 0 to 1
    eCutting := 30,   // 切割窗口：速比恒 1，bCutReq 置位 / Cutting window, ratio held 1, cut request active
    eSyncOut := 40    // 同步返回：速比 1→0 对称降回 / Sync-out, ratio ramping 1 back to 0
);
END_TYPE

(*==============================================================================
 * 功能块: FB_DL_FlyingSawSyncSeq
 * 调用约定: 每个扫描周期无条件调用一次；实例状态全部驻留于私有变量。
 * 调用示例: sawSeq(bEn := bLineRun, bStart := bBatchGo,
 *                  fMasterPos := fEncPos, fSyncLen := 120.0, fCutLen := 25.0);
 *          刀轴速度指令 = fEncVel × sawSeq.fRatio；bCutReq 触发剪切执行器，
 *          bCycleDone 作为计件脉冲送上层台账。
 * 组装说明: ① 本件为纯位置闭环序列件，主轴位置经 PRG_IoMapping 读入后
 *             引脚注入，本件零 %I/%Q 物理地址（红线 R2）；
 *           ② bCutReq 属请求级信号，剪切电磁阀驱动须在上层输出映射层
 *             复加安全联锁（与急停链 FB_DL_EmergencyStopChainDiag 合取）；
 *           ③ 多刀位并行时每刀独立实例，主轴位置引脚共享即可。
 *==============================================================================*)
FUNCTION_BLOCK FB_DL_FlyingSawSyncSeq
VAR_INPUT
    bEn        : BOOL := FALSE;        // 使能（FALSE 冻结回怠速）/ Enable, FALSE freezes to idle
    bStart     : BOOL := FALSE;        // 单周期启动沿输入 / One-cycle start trigger input
    fMasterPos : LREAL := 0.0;         // 同步轴位置 [mm]，序列时钟 / Master axis position [mm], the sequence clock
    fSyncLen   : LREAL := 100.0;       // 同步窗长度（切入=返回对称）[mm] / Sync window length, ramp-in equals ramp-out [mm]
    fCutLen    : LREAL := 20.0;        // 切割窗口长度（速比 1 区间）[mm] / Cutting window length at ratio 1 [mm]
END_VAR
VAR_OUTPUT
    bKnifeRun  : BOOL;                 // 刀轴运行使能输出 / Knife axis run enable output
    fRatio     : LREAL;                // 主从速比 [1]，刀速 = 主速 × 本值 / Master-to-knife velocity ratio [1]
    bCutReq    : BOOL;                 // 切割请求（速比 1 窗口内）[—] / Cut request inside the ratio-1 window
    bCycleDone : BOOL;                 // 单拍完成脉冲（本拍有效）[—] / Single-scan cycle-done pulse
    eState     : E_DL_FlyingSawState;  // 序列当前相位 / Current sequence phase
    uErrCode   : UDINT;                // 信息级码，0 = 无信息 / Info-level code, 0 = none
    bValid     : BOOL;                 // 输出有效标志（非有限拍为 FALSE）/ Outputs usable flag
END_VAR
VAR
    trigStart  : R_TRIG;               // 启动沿检测，每拍无条件刷新 / Start edge detector, refreshed every scan
    fAnchor    : LREAL;                // 切割锚点 [mm]，启动沿锁存为前方未来点（当前位置 + fSyncLen）/ Cut anchor [mm], latched ahead of the master (current position + fSyncLen)
    fLastPos   : LREAL;                // 主轴位置上拍快照 [mm]，防倒退闸用 / Master position last-scan snapshot [mm], reversal guard
    bEnEff     : BOOL;                 // 防御闸后的有效使能 / Effective enable after the defense gate
    _bDone     : BOOL;                 // 完成脉冲内部暂存（统一出口映射） / Done pulse internal stage, mapped at the unified outlet
END_VAR
VAR CONSTANT
    DL_FS_EPS  : LREAL := 1.0E-9;      // 浮点容差（窗长下限闸）[mm] / Float tolerance, window length floor [mm]
    DL_FS_INF  : LREAL := 1.7976931348623157E308; // LREAL 幅值上限 / LREAL magnitude ceiling
END_VAR

// ---- 段 1｜沿实例无条件刷新 + 单拍脉冲出口（两段式：置位在 CASE，映射在此）----
trigStart(CLK := bStart);              // 启动沿每拍刷新 / Start edge refreshed unconditionally
_bDone := FALSE;                       // 完成脉冲暂存先清零 / Done stage preset FALSE
bCutReq := FALSE;                      // 切割请求默认 FALSE（切割相内重置位）/ Cut request preset FALSE, re-raised in the cutting phase

// ---- 段 2｜输入防御与参数闸：非有限或参数退化 → 安全侧拒绝（信息级）----
IF (fMasterPos <> fMasterPos) OR (ABS(fMasterPos) > DL_FS_INF)
   OR (fSyncLen <> fSyncLen) OR (ABS(fSyncLen) > DL_FS_INF)
   OR (fCutLen <> fCutLen) OR (ABS(fCutLen) > DL_FS_INF) THEN
    bEnEff   := FALSE;                 // 非有限输入冻结使能 / Non-finite input freezes the enable
    eState   := eIdle;                 // 序列强制回怠速（安全侧）/ Sequence forced back to idle, safe side
    fAnchor  := 0.0;                   // 锚点清零防残留 / Anchor cleared against stale value
    uErrCode := 16#0004_08C0;          // 信息级：输入非有限 / Info: non-finite input
    bValid   := FALSE;                 // 输出不可用 / Outputs unusable
    RETURN;                            // 结构早退（输出保持确定值）/ early exit with deterministic outputs
END_IF
IF (fSyncLen <= DL_FS_EPS) OR (fCutLen <= DL_FS_EPS) THEN
    bEnEff   := FALSE;                 // 参数退化冻结使能 / Degenerated parameters freeze the enable
    eState   := eIdle;                 // 回怠速并留痕 / Back to idle with the code set
    uErrCode := 16#0004_08C0;          // 信息级：窗长参数非法 / Info: illegal window length
    bValid   := FALSE;                 // 输出不可用 / Outputs unusable
    RETURN;                            // 结构早退 / early exit
END_IF
bEnEff   := bEn;                       // 闸后有效使能 / Effective enable after the gate
uErrCode := 16#0000_0000;              // 信息码先清零 / Info code cleared first
bValid   := TRUE;                      // 防御通过输出可用 / Outputs usable after the gate

// ---- 段 3｜序列状态机（CASE 带 ELSE 非法态兜底；速比统一出口赋值）----
CASE eState OF
    E_DL_FlyingSawState.eIdle:         // 怠速相：等待启动沿
        fRatio := 0.0;                 // 速比零（安全侧）/ Ratio zero, safe side
        IF bEnEff AND trigStart.Q THEN
            fAnchor := fMasterPos + fSyncLen; // 锚点 = 当前位置 + 同步窗长（未来窗，切入区间落在主轴前方，R73）/ Anchor = current position + sync length, future window ahead of the master
            eState  := E_DL_FlyingSawState.eWait; // 进入待同步相 / Enter the waiting phase
        END_IF

    E_DL_FlyingSawState.eWait:         // 待同步相：等主轴进入同步窗
        fRatio := 0.0;                 // 未同步区间速比保持零 / Ratio held zero before the sync window
        IF NOT bEnEff THEN
            eState := E_DL_FlyingSawState.eIdle; // 撤使能中止 / Abort on disable
        ELSIF fMasterPos >= (fAnchor - fSyncLen) THEN
            eState := E_DL_FlyingSawState.eSyncIn; // 进入切入相 / Enter the ramp-in phase
        END_IF

    E_DL_FlyingSawState.eSyncIn:       // 切入相：速比 = 位置进度线性爬升
        fRatio := (fMasterPos - (fAnchor - fSyncLen)) / fSyncLen; // 进度比 [1]，分母已闸 / Progress ratio, denominator gated
        fRatio := MIN(MAX(fRatio, 0.0), 1.0);  // 速比双侧钳位 / Two-sided ratio clamp
        IF NOT bEnEff THEN
            eState := E_DL_FlyingSawState.eIdle;   // 撤使能中止 / Abort on disable
        ELSIF fMasterPos >= fAnchor THEN
            eState := E_DL_FlyingSawState.eCutting; // 到锚点进入切割相 / Reach the anchor, enter cutting
        END_IF

    E_DL_FlyingSawState.eCutting:      // 切割相：速比恒 1，切割请求置位
        fRatio  := 1.0;                // 完全同步 / Fully synchronized
        bCutReq := TRUE;               // 切割窗口声明 / Cut request declared
        IF NOT bEnEff THEN
            eState := E_DL_FlyingSawState.eIdle;   // 撤使能中止 / Abort on disable
        ELSIF fMasterPos >= (fAnchor + fCutLen) THEN
            eState := E_DL_FlyingSawState.eSyncOut; // 出切割窗进入返回相 / Leave the window, enter ramp-out
        END_IF

    E_DL_FlyingSawState.eSyncOut:      // 返回相：速比对称降回 0
        fRatio := 1.0 - (fMasterPos - (fAnchor + fCutLen)) / fSyncLen; // 对称进度比 [1] / Mirrored progress ratio
        fRatio := MIN(MAX(fRatio, 0.0), 1.0);  // 速比双侧钳位 / Two-sided ratio clamp
        IF NOT bEnEff THEN
            eState := E_DL_FlyingSawState.eIdle;   // 撤使能中止 / Abort on disable
        ELSIF fMasterPos >= (fAnchor + fCutLen + fSyncLen) THEN
            eState := E_DL_FlyingSawState.eIdle;   // 序列完成回怠速 / Sequence complete, back to idle
            _bDone := TRUE;                        // 完成脉冲内部置位（出口统一映射） / Done stage set, mapped at the outlet
        END_IF

    ELSE                               // 非法状态兜底（R21：CASE 必带 ELSE）
        eState  := E_DL_FlyingSawState.eIdle;      // 拦截非法值回怠速 / Catch illegal value back to idle
        fRatio  := 0.0;                // 速比归零（安全侧）/ Ratio zeroed, safe side
END_CASE

// ---- 段 4｜防倒退闸：活动相内主轴位置倒退 → 序列中止回怠速（安全侧）----
IF (eState = E_DL_FlyingSawState.eSyncIn)
   OR (eState = E_DL_FlyingSawState.eCutting)
   OR (eState = E_DL_FlyingSawState.eSyncOut) THEN
    IF fMasterPos < (fLastPos - DL_FS_EPS) THEN // 位置倒退超容差判方向反转 / Position regression beyond tolerance, reversal
        eState   := E_DL_FlyingSawState.eIdle;  // 序列中止回怠速 / Sequence aborted to idle
        fRatio   := 0.0;               // 速比归零（安全侧）/ Ratio zeroed, safe side
        uErrCode := 16#0004_08C0;      // 信息级：主轴方向反转中止（复用码 R90）/ Info: reversal abort, code reused
        bValid   := FALSE;             // 本拍输出不可信 / Outputs unusable this scan
    END_IF
END_IF
fLastPos := fMasterPos;                // 位置快照滚存（闸后统一写）/ Snapshot rolled forward after the gate

// ---- 段 5｜统一出口：完成脉冲单拍映射 + 速比安全兜底 ----
bCycleDone := _bDone;                  // 完成脉冲本拍有效 / Done pulse valid this scan
bKnifeRun  := bEn AND (eState <> E_DL_FlyingSawState.eIdle); // 运行使能随相位 / Run enable follows the phase
END_FUNCTION_BLOCK

(* ---- FB_DL_GantryCraneAnchoringSeq.st ---- *)
(*
 * FB_DL_GantryCraneAnchoringSeq | C4 | DL_Motion
 * 功能：大车自动锚定与防风防滑序列（风速分级→减速→夹轨→锚定→解除）；每相独立使能出口 + 独立 TON 超时，超时回 FAULT 并回退全部命令       单位：rWindMs [m/s]、rTimeoutS [s]、nFaultCode [INT 码位]
 * 工况边界：工作状态风速 0~40 m/s（GB/T 3811 分级：<13.8 正常 / 13.8~20 降速 / 20~25 停工夹轨锚定 / >25 直接锚定）；rTimeoutS 须 >0；解除仅当风速 <13.8、xRelease 有效且锚定驻留已满一个超时窗；全速许可须在 IDLE 稳定驻留满一个超时窗才恢复；风速 NaN/±Inf 一律按最不利(锚定侧)处理；IDLE/WIND_WARN/DECEL/ANCHORED 的 TON 为监督/驻留定时（驻留超时只置信息码 9106，绝不升级为锚定），CLAMPING/ANCHORING/RELEASING 的 TON 为故障超时（码表见下）；xEnable=FALSE 时两路输出回落失电安全侧（夹轨/锚定销弹簧夹紧型），但**不改变相位**
 * 代数值回代：rWindMs=22.0 → DECEL→CLAMPING→ANCHORED（20~25 区间）；rWindMs=26.0 → 直跳 ANCHORING；rWindMs=8.0 且 xRelease=TRUE → RELEASING→IDLE（与 spec 分级回代一致）
 * 开源溯源：clean-room 自研，未复制任何第三方代码（无外部来源）
 *)
(*
 * 码位总账（本件故障码全清单，逐条在实现分支中可到达；故障级锁存回放）：
 * 9101 夹轨超时 / 9102 锚定超时 / 9103 解除超时 / 9104 风速越限解除被拒 / 9105 入参非有限或状态机兜底 / 9106 降速相驻留超时（信息级，不置故障）——故障锁存，清除沿 = xEnable 下降沿（仅下降沿，不用电平）
 *)

TYPE E_DL_GcAnchorPhase :
(
    IDLE      := 0,      // 待机，允许行车，无夹轨无锚定命令 | idle, travelling permitted, no clamp and no anchor command
    WIND_WARN := 10,     // 降速相，风速 13.8~20，允许低速行车 | derated phase, wind 13.8 to 20, slow travel permitted
    DECEL     := 20,     // 减速停车相，风速 20~25，撤销行车许可 | deceleration phase, wind 20 to 25, travel permit withdrawn
    CLAMPING  := 30,     // 夹轨相，等夹轨到位反馈 | clamping phase, waiting for the rail clamp feedback
    ANCHORING := 40,     // 锚定相，等锚定到位反馈 | anchoring phase, waiting for the anchor feedback
    ANCHORED  := 50,     // 已锚定稳态，全部防风机构到位 | anchored steady state, all wind devices engaged
    RELEASING := 60,     // 解除相，等夹轨与锚定同时松开 | releasing phase, waiting for clamp and anchor to retract
    FAULT     := 90      // 故障相，全部命令回退为 FALSE，码位锁存 | fault phase, every command reverts to FALSE, the code is latched
);
END_TYPE

FUNCTION_BLOCK FB_DL_GantryCraneAnchoringSeq
VAR_INPUT
    xEnable      : BOOL;             // 序列总使能（下降沿兼作故障复位沿）| sequence enable, its falling edge also resets a latched fault
    xRelease     : BOOL;             // 解除请求，仅风速 <13.8 时被接受 | release request, accepted only when the wind is below 13.8
    rWindMs      : REAL;             // 实测风速（3 s 均值）| measured wind speed, 3 s mean [m/s]
    xRailClampFb : BOOL;             // 夹轨到位反馈 | rail clamp engaged feedback
    xAnchorFb    : BOOL;             // 锚定销到位反馈 | anchor pin engaged feedback
    rTimeoutS    : REAL := 20.0;     // 每相超时设定 | per-phase timeout setting [s]
END_VAR
VAR_OUTPUT
    xClampCmd       : BOOL;          // 夹轨命令（仅 CLAMPING/ANCHORING/ANCHORED 为 TRUE）| rail clamp command, TRUE in CLAMPING, ANCHORING and ANCHORED only
    xAnchorCmd      : BOOL;          // 锚定命令（仅 ANCHORING/ANCHORED 为 TRUE）| anchor command, TRUE in ANCHORING and ANCHORED only
    ePhase          : E_DL_GcAnchorPhase;  // 当前相 | current phase
    xPermitTravel   : BOOL;          // 行车许可（仅 IDLE 与 WIND_WARN 为 TRUE）| travel permit, TRUE in IDLE and WIND_WARN only
    xPermitFullSpeed: BOOL;          // 全速许可（仅 IDLE 为 TRUE）| full speed permit, TRUE in IDLE only
    xFault          : BOOL;          // 故障标志（故障级码才置位）| fault flag, raised by fault-class codes only
    nFaultCode      : INT;           // 故障码，锁存至复位沿 | fault code, latched until the reset edge
END_VAR
VAR
    tonIdle     : TON;               // IDLE 相监督定时器 | supervision timer of the IDLE phase
    tonWarn     : TON;               // WIND_WARN 相驻留定时器 | dwell timer of the WIND_WARN phase
    tonDecel    : TON;               // DECEL 相减速驻留定时器 | deceleration dwell timer of the DECEL phase
    tonClampTmo : TON;               // CLAMPING 相故障超时定时器 | fault timeout of the CLAMPING phase
    tonAnchorTmo: TON;               // ANCHORING 相故障超时定时器 | fault timeout of the ANCHORING phase
    tonAnchored : TON;               // ANCHORED 相监督定时器 | supervision timer of the ANCHORED phase
    tonReleaseTmo: TON;              // RELEASING 相故障超时定时器 | fault timeout of the RELEASING phase
    fbEnableFall: F_TRIG;            // xEnable 下降沿检测（故障复位沿）| falling edge of xEnable, the fault reset edge
    xFinWind    : BOOL;              // 风速有限性 | wind speed is finite
    xWindBad    : BOOL;              // 风速非有限或超量程 | wind speed non-finite or out of range
    xParamOk    : BOOL;              // 超时参数合法（有限且 >0）| timeout parameter is legal, finite and positive
    nTmoMs      : UDINT := 20000;    // 超时毫秒数（REAL→UDINT 标准转换，缺省值防首拍 PT=0）| timeout in milliseconds with a default preventing a zero PT on the first scan
    nDecelMs    : UDINT := 3000;     // 减速驻留毫秒数 | deceleration dwell in milliseconds
    rWindChk    : REAL;              // 判定用风速（非有限时置最不利值）| wind value used for grading, forced to the worst case when non-finite
    nCodeLatch  : INT;               // 故障码锁存副本 | latched copy of the fault code
END_VAR
VAR CONSTANT
    DL_GCA_WIND_DERATE : REAL := 13.8;   // 降速风速阈 | derating wind threshold [m/s]
    DL_GCA_WIND_STOP   : REAL := 20.0;   // 停工夹轨风速阈 | stop and clamp wind threshold [m/s]
    DL_GCA_WIND_ANCHOR : REAL := 25.0;   // 强制锚定风速阈 | mandatory anchoring wind threshold [m/s]
    DL_GCA_WIND_MAX    : REAL := 40.0;   // 风速量程上限 | upper wind range limit [m/s]
    DL_GCA_DECEL_S     : REAL := 3.0;    // 减速驻留时间（变频器斜坡）| deceleration dwell matching the drive ramp [s]
    DL_GCA_C_WIND_OVER : INT := 9104;    // 风速越限解除被拒 | release refused because the wind is over limit
    DL_GCA_C_CLAMP_TMO : INT := 9101;    // 夹轨超时 | rail clamp timeout
    DL_GCA_C_ANCH_TMO  : INT := 9102;    // 锚定超时 | anchoring timeout
    DL_GCA_C_REL_TMO   : INT := 9103;    // 解除超时 | releasing timeout
    DL_GCA_C_BAD       : INT := 9105;    // 入参非有限或状态机兜底 | non-finite input or state machine fallback
    DL_GCA_I_WARN_DWELL : INT := 9106;   // 信息级：降速相驻留超时（不置 xFault）| info level, derated phase dwell expired
END_VAR

// 段1｜参数与采样门禁（先判后用：所有 REAL→UDINT 换算在闸后进行；换算结果供段2 定时器使用）
xParamOk := (rTimeoutS = rTimeoutS) AND ((rTimeoutS - rTimeoutS) = 0.0) AND (rTimeoutS > 0.0);
xFinWind := (rWindMs = rWindMs) AND ((rWindMs - rWindMs) = 0.0);
xWindBad := (NOT xFinWind) OR (rWindMs < 0.0) OR (rWindMs > DL_GCA_WIND_MAX);
IF xWindBad THEN
    rWindChk := DL_GCA_WIND_MAX;     // 风速不可信一律按最不利（锚定侧）分级 | an untrusted wind value is graded at the worst case
ELSE
    rWindChk := rWindMs;
END_IF
IF NOT xParamOk THEN
    nTmoMs := 20000;                 // 参数非法时的保守超时 | conservative timeout when the parameter is illegal
    nDecelMs := 3000;
ELSE
    nTmoMs := REAL_TO_UDINT(rTimeoutS * 1000.0);
    nDecelMs := REAL_TO_UDINT(DL_GCA_DECEL_S * 1000.0);
END_IF

// 段2｜七只定时器 + 一只边沿实例无条件周期刷新（R7：严禁放入 IF/CASE，一相一只实例不跨相复用）
// PT 取自段1 已换算的毫秒值；声明缺省值保证首拍 PT 不为 0，不会出现首拍即 Q=TRUE 的假超时
tonIdle(IN := (ePhase = E_DL_GcAnchorPhase.IDLE) AND xEnable, PT := UDINT_TO_TIME(nTmoMs));
tonWarn(IN := ePhase = E_DL_GcAnchorPhase.WIND_WARN, PT := UDINT_TO_TIME(nTmoMs));
tonDecel(IN := ePhase = E_DL_GcAnchorPhase.DECEL, PT := UDINT_TO_TIME(nDecelMs));
tonClampTmo(IN := ePhase = E_DL_GcAnchorPhase.CLAMPING, PT := UDINT_TO_TIME(nTmoMs));
tonAnchorTmo(IN := ePhase = E_DL_GcAnchorPhase.ANCHORING, PT := UDINT_TO_TIME(nTmoMs));
tonAnchored(IN := ePhase = E_DL_GcAnchorPhase.ANCHORED, PT := UDINT_TO_TIME(nTmoMs));
tonReleaseTmo(IN := ePhase = E_DL_GcAnchorPhase.RELEASING, PT := UDINT_TO_TIME(nTmoMs));
fbEnableFall(CLK := xEnable);

// 段3｜输出预置（出口唯一预置点，CASE 内只置位，绝不在其后无条件清零）
xClampCmd := FALSE;
xAnchorCmd := FALSE;
xPermitTravel := FALSE;
xPermitFullSpeed := FALSE;
xFault := FALSE;
nFaultCode := 0;

// 段4｜主状态机（ENUM + CASE，含 ELSE 兜底）
CASE ePhase OF
E_DL_GcAnchorPhase.IDLE:
    // 拍 N 进入：IDLE，夹轨与锚定均复位，行车许可有效
    xPermitTravel := TRUE;                                   // 本拍行为：行车许可（降速以上即撤）| this scan: travel permitted
    xPermitFullSpeed := tonIdle.Q;                           // 全速许可须在 IDLE 稳定驻留满一个超时窗（风速持续低于降速阈）| full speed only after a stable dwell
    IF xWindBad THEN
        ePhase := E_DL_GcAnchorPhase.ANCHORING;              // 风速不可信：跳级直锚（安全侧）| untrusted wind, anchor at once
    ELSIF rWindChk > DL_GCA_WIND_ANCHOR THEN
        ePhase := E_DL_GcAnchorPhase.ANCHORING;              // >25：直接锚定 | above 25, anchor directly
    ELSIF rWindChk > DL_GCA_WIND_STOP THEN
        ePhase := E_DL_GcAnchorPhase.DECEL;                  // 20~25：先减速再夹轨锚定 | 20 to 25, decelerate then clamp and anchor
    ELSIF rWindChk >= DL_GCA_WIND_DERATE THEN
        ePhase := E_DL_GcAnchorPhase.WIND_WARN;              // 13.8~20：降速 | 13.8 to 20, derate
    END_IF
    // 拍 N+1：若进 ANCHORING/DECEL，本拍命令仍全 FALSE（命令在目标相置位）

E_DL_GcAnchorPhase.WIND_WARN:
    // 拍 N 进入：降速相，行车许可保留、全速许可撤销
    xPermitTravel := TRUE;                                   // 本拍行为：仅保留降速行车许可 | this scan: derated travel only
    xPermitFullSpeed := FALSE;
    IF rWindChk > DL_GCA_WIND_STOP THEN
        ePhase := E_DL_GcAnchorPhase.DECEL;                  // 升过 20：转减速 | above 20, go to deceleration
    ELSIF rWindChk < DL_GCA_WIND_DERATE - 1.0 THEN
        ePhase := E_DL_GcAnchorPhase.IDLE;                   // 回落 1 m/s 滞环后恢复全速（须先于驻留判定，否则 Q 恒真致本分支永不可达）| hysteresis first, otherwise tonWarn.Q latches and blocks it
    ELSIF tonWarn.Q THEN
        nFaultCode := DL_GCA_I_WARN_DWELL;                   // 降速相驻留超时：仅置信息码，不升级为锚定（13.8~20 m/s 属降速作业区，GB/T 3811）| dwell expired, informational only, no escalation
    END_IF

E_DL_GcAnchorPhase.DECEL:
    // 拍 N 进入：减速停车，行车许可撤销，夹轨命令尚未给出
    IF tonDecel.Q THEN
        ePhase := E_DL_GcAnchorPhase.CLAMPING;               // 本拍行为：减速完成转夹轨 | deceleration done, go to clamping
    ELSIF rWindChk > DL_GCA_WIND_ANCHOR THEN
        ePhase := E_DL_GcAnchorPhase.ANCHORING;              // 超 25：跳过夹轨直锚 | above 25, skip clamping and anchor
    END_IF

E_DL_GcAnchorPhase.CLAMPING:
    // 拍 N 进入：夹轨命令置位（段5），等夹轨到位反馈
    IF xRailClampFb THEN
        ePhase := E_DL_GcAnchorPhase.ANCHORING;              // 本拍行为：夹轨到位转锚定 | clamp engaged, go to anchoring
    ELSIF tonClampTmo.Q THEN
        nCodeLatch := DL_GCA_C_CLAMP_TMO;                    // 夹轨超时：锁存 9101 | clamp timeout, latch 9101
        xFault := TRUE;
        nFaultCode := DL_GCA_C_CLAMP_TMO;
        ePhase := E_DL_GcAnchorPhase.FAULT;
    END_IF

E_DL_GcAnchorPhase.ANCHORING:
    // 拍 N 进入：夹轨 + 锚定命令同时置位（段5），等锚定销到位
    IF xAnchorFb AND xRailClampFb THEN
        ePhase := E_DL_GcAnchorPhase.ANCHORED;               // 本拍行为：双到位转锚定稳态 | both engaged, go to the anchored steady state
    ELSIF tonAnchorTmo.Q THEN
        nCodeLatch := DL_GCA_C_ANCH_TMO;                     // 锚定超时：锁存 9102 | anchoring timeout, latch 9102
        xFault := TRUE;
        nFaultCode := DL_GCA_C_ANCH_TMO;
        ePhase := E_DL_GcAnchorPhase.FAULT;
    END_IF

E_DL_GcAnchorPhase.ANCHORED:
    // 拍 N 进入：稳态锚定，行车许可全撤
    IF (NOT xAnchorFb) OR (NOT xRailClampFb) THEN
        ePhase := E_DL_GcAnchorPhase.ANCHORING;              // 反馈丢失：回锚定相重试（超时由 9102 兜底）| feedback lost, retry anchoring
    ELSIF xRelease AND tonAnchored.Q AND (rWindChk < DL_GCA_WIND_DERATE) THEN
        ePhase := E_DL_GcAnchorPhase.RELEASING;              // 本拍行为：锚定驻留满足且风速达标，转解除相 | dwell satisfied and wind low, go to releasing
    ELSIF xRelease AND (rWindChk >= DL_GCA_WIND_DERATE) THEN
        nFaultCode := DL_GCA_C_WIND_OVER;                    // 信息级：风速越限解除被拒（不置 xFault）| info: release refused because of the wind
    END_IF

E_DL_GcAnchorPhase.RELEASING:
    // 拍 N 进入：解除相，夹轨与锚定命令均撤销（段5）
    IF (NOT xAnchorFb) AND (NOT xRailClampFb) THEN
        ePhase := E_DL_GcAnchorPhase.IDLE;                   // 本拍行为：双松开转待机 | both retracted, back to idle
    ELSIF rWindChk >= DL_GCA_WIND_DERATE THEN
        nCodeLatch := DL_GCA_C_WIND_OVER;                    // 解除中风速回升：回锚定并锁 9104 | wind rose during release, re-anchor and latch 9104
        xFault := TRUE;
        nFaultCode := DL_GCA_C_WIND_OVER;
        ePhase := E_DL_GcAnchorPhase.FAULT;
    ELSIF tonReleaseTmo.Q THEN
        nCodeLatch := DL_GCA_C_REL_TMO;                      // 解除超时：锁存 9103 | releasing timeout, latch 9103
        xFault := TRUE;
        nFaultCode := DL_GCA_C_REL_TMO;
        ePhase := E_DL_GcAnchorPhase.FAULT;
    END_IF

E_DL_GcAnchorPhase.FAULT:
    // 拍 N 进入：故障相，全部命令回退 FALSE，码位锁存重发布
    xClampCmd := FALSE;                                      // 本拍行为：夹轨命令回退 | this scan: clamp command reverted
    xAnchorCmd := FALSE;                                     // 本拍行为：锚定命令回退 | this scan: anchor command reverted
    xFault := TRUE;
    nFaultCode := nCodeLatch;                                // 锁存回放，不在故障相按当下输入重推断 | republish the latch instead of re-inferring
    IF fbEnableFall.Q THEN
        nCodeLatch := 0;                                     // 清除边：仅 xEnable 下降沿（电平清除会导致故障每拍被清、锚定销周期性重击）| clear on the falling edge only
        ePhase := E_DL_GcAnchorPhase.IDLE;
    END_IF

ELSE
    // 非法状态兜底：绝不停在未知相
    nCodeLatch := DL_GCA_C_BAD;                              // 兜底锁存 9105 | fallback latches 9105
    xFault := TRUE;
    nFaultCode := DL_GCA_C_BAD;
    xClampCmd := FALSE;
    xAnchorCmd := FALSE;
    ePhase := E_DL_GcAnchorPhase.FAULT;
END_CASE

// 段5｜每相独立使能出口（故障与兜底相不置任何命令，天然强制 FALSE）
CASE ePhase OF
E_DL_GcAnchorPhase.CLAMPING:
    xClampCmd := TRUE;                                       // 夹轨相独立使能出口 | independent enable output of the clamping phase
E_DL_GcAnchorPhase.ANCHORING:
    xClampCmd := TRUE;                                       // 锚定相：夹轨保持 | anchoring, keep the clamp
    xAnchorCmd := TRUE;                                      // 锚定相独立使能出口 | independent enable output of the anchoring phase
E_DL_GcAnchorPhase.ANCHORED:
    xClampCmd := TRUE;                                       // 锚定稳态：夹轨保持 | anchored, keep the clamp
    xAnchorCmd := TRUE;                                      // 锚定稳态：锚定保持 | anchored, keep the anchor
E_DL_GcAnchorPhase.RELEASING:
    xClampCmd := FALSE;                                      // 解除相：夹轨撤销 | releasing, clamp retracted
    xAnchorCmd := FALSE;                                     // 解除相：锚定撤销 | releasing, anchor retracted
ELSE
    xClampCmd := FALSE;                                      // 其余相（含 FAULT）：命令强制 FALSE | all other phases force FALSE
    xAnchorCmd := FALSE;
END_CASE

// 段5b｜总使能门（R750）：未使能不得驱动夹轨/锚定机构
// 本件两路输出定义为失电即动作型（夹轨/锚定销弹簧夹紧、液压释放），FALSE 即安全侧，故使能撤销时回落 FALSE 是安全的
IF NOT xEnable THEN
    xClampCmd := FALSE;                                      // 未使能：夹轨命令回落失电安全侧 | disabled, clamp command falls back to the de-energised safe side
    xAnchorCmd := FALSE;                                     // 未使能：锚定命令回落失电安全侧 | disabled, anchor command falls back to the de-energised safe side
END_IF

// 段6｜出口汇总：非 IDLE/WIND_WARN 一律撤销行车许可；故障相已由段3预置为 FALSE
IF (ePhase <> E_DL_GcAnchorPhase.IDLE) AND (ePhase <> E_DL_GcAnchorPhase.WIND_WARN) THEN
    xPermitTravel := FALSE;                                  // 非行车相撤销许可 | non-travel phases withdraw the permit
    xPermitFullSpeed := FALSE;
END_IF
IF xWindBad THEN
    xPermitTravel := FALSE;                                  // 风速不可信：许可也撤 | untrusted wind withdraws the permit as well
    xPermitFullSpeed := FALSE;
END_IF
IF NOT xEnable THEN
    xPermitTravel := FALSE;                                  // 序列未使能：不给行车许可（R191 名实双出口）| sequence disabled, no travel permit
    xPermitFullSpeed := FALSE;
END_IF
END_FUNCTION_BLOCK

(* ---- FB_DL_GantryDualDriveTorqueBalance.st ---- *)
(*
    FB_DL_GantryDualDriveTorqueBalance —— 龙门双驱转矩失衡评估与从动侧偏置自适应
    ------------------------------------------------------------------
    组件名    : FB_DL_GantryDualDriveTorqueBalance
    分类      : DL_Motion / Dual-Drive Balance（双驱转矩均衡）
    一句话功能: 在线评估龙门双驱的转矩失衡，带死区按周期步进调整从动侧转矩偏置，
                失衡恶化时输出降速比例保护机械。
    复杂度    : C3
    版本      : v1.0.0
    开源溯源  : 无（clean-room 自研，未借鉴任何开源实现）
    平台      : 纯 IEC 61131-3（TON / R_TRIG / ABS 标准库），目标编译器 RuSTy 1.0.8，
                兼容 CODESYS 3.5 / TwinCAT 3 / 汇川 InoProShop / Machine Expert；
                无 PROPERTY、无 VLA、无 FOR..DOWNTO、无 AS 类方言
    ------------------------------------------------------------------
    功能说明  : ① 失衡度 fImbalancePct = ABS(fTorqueMasterPct − fTorqueSlavePct)，单位 %；
                ② 死区：失衡 ≤ fBalanceTolPct 时完全不调整偏置（防积分漂移抖动），
                   且 bBalanced := TRUE；
                ③ 调整：失衡 > 死区且处 eBiasAdj 相时，每 tBiasPeriodMs（TON 自复位，R188）
                   按 fBiasStepPct 朝「减小失衡」的方向步进一次 fBiasOutPct，并钳位在
                   ±fMaxBiasPct；方向约定：主轴转矩大（从动侧出力不足）→ 偏置加，反之偏置减；
                ④ 降额：失衡 > fBalanceTolPct × fDerateRatio → eDerate，fSpeedScalePct 从 100
                   线性降到 50 并饱和；恢复带滞回 fThDerate − DL_GB_HYS_PCT，防临界抖动；
                ⑤ 安全默认：bReset 上升沿与 eFault 相内 fBiasOutPct 一律清 0（不带偏置上电）；
                ⑥ 转矩读数非有限（NaN / ±Inf / 超幅值域）→ eFault，fSpeedScalePct := 0。
    量纲链    : fTorqueMasterPct [%] − fTorqueSlavePct [%] → 失衡度 fImbalancePct [%]（同类量相减）；
                fBalanceTolPct [%] × fDerateRatio [-] → 降额阈值 fThDerate [%]（比例无因次）；
                (fImbalancePct − fThDerate) [%] ÷ fThDerate [%] → _fRto [-]（% ÷ % 无因次）；
                fSpeedScalePct = 100 [%] − (100 − 50)[%] × _fRto [-] → [%]；
                fBiasStepPct [%] 逐拍累加到 fBiasOutPct [%]，钳位界 ±fMaxBiasPct [%]。
                全程无「温度、时间、角度进入转矩加法链」，量纲链逐段闭合。
    状态机    : eIdle(0) --使能且组态合法且数据有限--> eBalance(10)
                eBalance --失衡 > 死区--> eBiasAdj(20)；--失衡 > 降额阈值--> eDerate(30)
                eBiasAdj --失衡回到死区内--> eBalance（偏置保持）；--失衡 > 降额阈值--> eDerate
                eDerate --失衡 ≤ 降额阈值 − DL_GB_HYS_PCT--> 回到 eBalance 或 eBiasAdj
                任意相 --失能--> eIdle；--数据非有限或组态非法--> eFault(90)
                eFault 的唯一解除路径 = bReset 上升沿（见段 8 与复位作用域声明）
    失能语义  : bEnable = FALSE → eIdle，fBiasOutPct 清 0、fSpeedScalePct 清 0（安全侧：不带偏置、
                不发放行），不冻结末次偏置 —— 双驱偏置在无人监控时保持是有害的（R191 显式声明）。
    复位作用域: bReset 上升沿①清 _bFaultLatch / _bBadIn / _bCfgBad；②fBiasOutPct 清 0 且
                _fBias 清 0（偏置不得跨复位继承）；③迁相回 eIdle；④不清 _fImb（下一拍重算）。
    防御口径  : NaN 用自反 f<>f；±Inf 用 (f−f)<>(f−f)；另设幅值域闸 ABS(f) > 1.0E30。
                除法前先判零：降额归一的分母 fThDerate 与 DL_GB_EPS 比较后才做除法，组态闸另
                强制 fBalanceTolPct > DL_GB_EPS 且 fDerateRatio > 1.0，使分母结构性为正。
                周期调整 TON 的 IN 由自身 Q 取反驱动（IN := NOT tonBias.Q ...），不依赖外部沿（R188）。
    规格补充  : 按 R190 归因唯一补充 bCfgErr / bDataErr 两个诊断位，使两条故障成因各自可观测。
    码位说明  : 本件按零码位范式交付，不分配 16# 事件码；失衡、降额与故障一律经
                eState / bBalanced / bFaultOut / bCfgErr / bDataErr 组合观测。
    修订记录  : 2026-11-24 v1.0.0 首次入库（R87 批 · #4）
*)
TYPE E_DL_BalanceState :
(
    eIdle    := 0,    // 空闲：未使能，偏置与放行均清 0 | idle, disabled, bias and release both zeroed
    eBalance := 10,   // 均衡：失衡在死区内，偏置保持不动 | balanced, imbalance inside the dead band, bias held
    eBiasAdj := 20,   // 偏置调整：按周期步进偏置以减小失衡 | bias adjustment, stepped once per period
    eDerate  := 30,   // 降额：失衡超降额阈值，输出降速比例 < 100 | derate, speed scale below 100
    eFault   := 90    // 故障：读数非有限或组态非法，锁存至复位沿 | fault latched until the reset edge
);
END_TYPE

FUNCTION_BLOCK FB_DL_GantryDualDriveTorqueBalance
VAR_INPUT
    bEnable          : BOOL;                      // 使能电平，TRUE = 允许评估与调整 | enable level, TRUE = evaluation and adjustment active
    bReset           : BOOL;                      // 复位请求，上升沿生效 | reset request, rising-edge active
    fTorqueMasterPct : REAL;                      // 主轴转矩百分比 [%]，可为负（回馈）| master torque [%], negative on regen
    fTorqueSlavePct  : REAL;                      // 从动轴转矩百分比 [%] | slave torque [%]
    fBalanceTolPct   : REAL := 5.0;               // 失衡死区（容差）[%]，须为正 | imbalance dead band [%]
    fMaxBiasPct      : REAL := 10.0;              // 偏置钳位上限 [%]，须为正 | bias clamp magnitude [%]
    fDerateRatio     : REAL := 3.0;               // 降额阈值相对死区的倍数 [-]，须 > 1 | derate threshold as a multiple of the band
    fBiasStepPct     : REAL := 0.5;               // 每周期偏置步长 [%]，须为正 | bias step per period [%]
    tBiasPeriodMs    : TIME := T#500MS;           // 偏置步进周期 [ms] | bias step period [ms]
END_VAR
VAR_OUTPUT
    eState           : E_DL_BalanceState;         // 主状态，供 HMI 与联锁使用 | main state for HMI and interlocks
    fImbalancePct    : REAL;                      // 本拍失衡度 [%] | imbalance this scan [%]
    fBiasOutPct      : REAL;                      // 从动侧转矩偏置指令 [%]，正 = 增加从动侧出力 | slave torque bias [%]
    fSpeedScalePct   : REAL;                      // 派生速度比例指令 [%]，100 = 不限速 | derived speed scale [%]
    bBalanced        : BOOL;                      // 失衡在死区内 | imbalance inside the dead band
    bFaultOut        : BOOL;                      // 故障汇总位 | fault aggregate
    bCfgErr          : BOOL;                      // 组态非法诊断位（归因唯一，R190）| bad-configuration flag
    bDataErr         : BOOL;                      // 数据非有限诊断位（归因唯一，R190）| non-finite data flag
END_VAR
VAR
    rtReset          : R_TRIG;                    // 复位上升沿实例，每拍无条件刷新 | reset rising-edge instance
    tonBias          : TON;                       // 偏置步进周期计时，自复位，每拍无条件刷新 | bias step period timer
    _eState          : E_DL_BalanceState := E_DL_BalanceState.eIdle; // 状态机内部当前态 | internal current state
    _bInit           : BOOL := TRUE;              // 首扫初始化标志，含偏置积分状态 | first-scan init flag
    _bResetLatch     : BOOL := FALSE;             // 复位沿锁存量，本拍末清除 | reset-edge latch, cleared at scan end
    _bFaultLatch     : BOOL := FALSE;             // 故障锁存位 | fault latch
    _bBadIn          : BOOL := FALSE;             // 数据非有限成因位 | non-finite data cause
    _bCfgBad         : BOOL := FALSE;             // 组态非法成因位 | bad configuration cause
    _fBias           : REAL := 0.0;               // 偏置累积值 [%] | accumulated bias [%]
    _fImb           : REAL := 0.0;                // 本拍失衡度 [%] | imbalance this scan [%]
    _fThDerate       : REAL := 0.0;               // 本拍降额阈值 [%] | derate threshold this scan [%]
    _fThRecover      : REAL := 0.0;               // 本拍降额恢复阈值 [%] | derate recovery threshold this scan [%]
    _fDen            : REAL := 0.0;               // 降额归一除子 [%] | derate normalisation divisor [%]
    _fRto            : REAL := 0.0;               // 降额带内归一比例 [0..1] | normalised ratio inside the derate band
END_VAR
VAR CONSTANT
    DL_GB_EPS        : REAL := 1.0E-6;            // 浮点判零容差 [%] | float zero tolerance [%]
    DL_GB_MAG_MAX    : REAL := 1.0E30;            // 有限幅值域闸上限 [%] | magnitude domain bound [%]
    DL_GB_SCALE_FULL : REAL := 100.0;             // 满速比例 [%] | full speed scale [%]
    DL_GB_SCALE_MIN  : REAL := 50.0;              // 降额最低速度比例 [%] | minimum derated speed scale [%]
    DL_GB_HYS_PCT    : REAL := 2.0;               // 降额恢复滞回带 [%] | derate release hysteresis [%]
    DL_GB_RATIO_MIN  : REAL := 1.0;               // 降额倍数的下界 [-]（须严格大于该值）| lower bound of the derate multiple
END_VAR

METHOD ClampBias : REAL
(*
    偏置钳位：把偏置钳到 ±fMaxBiasPct（调用方保证 fMaxBiasPct > 0 且有限）。纯函数，无跨拍状态。
    Clamp the bias to plus or minus the configured magnitude; the caller guarantees a positive finite limit.
*)
VAR_INPUT
    fIn   : REAL;                                 // 待钳偏置 [%] | bias to clamp [%]
    fLimit: REAL;                                 // 钳位界（正数）[%] | clamp magnitude, positive [%]
END_VAR
ClampBias := fIn;                                 // 直通后按两侧硬界饱和 | straight-through, saturated below
IF ClampBias > fLimit THEN
    ClampBias := fLimit;                          // 正向钳到 +界 [%] | clamp to the positive limit
END_IF
IF ClampBias < (0.0 - fLimit) THEN
    ClampBias := 0.0 - fLimit;                    // 负向钳到 −界 [%] | clamp to the negative limit
END_IF
END_METHOD

// 段 1｜输出预置与首扫初始化（含偏置积分状态，故必须有 _bInit，R310）
// segment 1, output presets and first-scan initialisation; the bias integrator requires _bInit
fSpeedScalePct := 0.0;                             // 预置速度比例 0 [%]，放行默认撤销 | preset zero speed scale
bBalanced := FALSE;                                // 预置非均衡 | preset not balanced
fBiasOutPct := 0.0;                                // 预置偏置 0 [%] | preset zero bias
_bBadIn := FALSE;                                  // 预置数据有限 | preset finite data
_bCfgBad := FALSE;                                 // 预置组态合法 | preset legal configuration
IF _bInit THEN
    _bInit := FALSE;                               // 首扫只执行一次 | runs once on the first scan
    _eState := E_DL_BalanceState.eIdle;            // 首扫状态回空闲相 | initialise the state
    _fBias := 0.0;                                 // 首扫偏置归零 [%]，不带偏置上电 | initial bias [%]
END_IF

// 段 2｜非有限闸：NaN 自反 + Inf 自减 + 幅值域，逐个浮点入参枚举（R4 / R151 / R272）
// segment 2, non-finite gate over every REAL input: NaN self-reflexive, Inf by self-subtraction, magnitude bound
IF (fTorqueMasterPct <> fTorqueMasterPct) OR ((fTorqueMasterPct - fTorqueMasterPct) <> (fTorqueMasterPct - fTorqueMasterPct)) THEN
    _bBadIn := TRUE;                               // 主轴转矩 NaN 或 ±Inf | master torque NaN or infinity
END_IF
IF ABS(fTorqueMasterPct) > DL_GB_MAG_MAX THEN
    _bBadIn := TRUE;                               // 主轴转矩超幅值域 | master torque beyond the magnitude domain
END_IF
IF (fTorqueSlavePct <> fTorqueSlavePct) OR ((fTorqueSlavePct - fTorqueSlavePct) <> (fTorqueSlavePct - fTorqueSlavePct)) THEN
    _bBadIn := TRUE;                               // 从动轴转矩 NaN 或 ±Inf | slave torque NaN or infinity
END_IF
IF ABS(fTorqueSlavePct) > DL_GB_MAG_MAX THEN
    _bBadIn := TRUE;                               // 从动轴转矩超幅值域 | slave torque beyond the magnitude domain
END_IF
IF (fBalanceTolPct <> fBalanceTolPct) OR ((fBalanceTolPct - fBalanceTolPct) <> (fBalanceTolPct - fBalanceTolPct)) THEN
    _bBadIn := TRUE;                               // 死区 NaN 或 ±Inf | dead band NaN or infinity
END_IF
IF (fMaxBiasPct <> fMaxBiasPct) OR ((fMaxBiasPct - fMaxBiasPct) <> (fMaxBiasPct - fMaxBiasPct)) THEN
    _bBadIn := TRUE;                               // 偏置上限 NaN 或 ±Inf | bias limit NaN or infinity
END_IF
IF (fDerateRatio <> fDerateRatio) OR ((fDerateRatio - fDerateRatio) <> (fDerateRatio - fDerateRatio)) THEN
    _bBadIn := TRUE;                               // 降额倍数 NaN 或 ±Inf | derate multiple NaN or infinity
END_IF
IF (fBiasStepPct <> fBiasStepPct) OR ((fBiasStepPct - fBiasStepPct) <> (fBiasStepPct - fBiasStepPct)) THEN
    _bBadIn := TRUE;                               // 步长 NaN 或 ±Inf | bias step NaN or infinity
END_IF
IF ABS(fBalanceTolPct) > DL_GB_MAG_MAX THEN
    _bBadIn := TRUE;                               // 死区超幅值域 | dead band beyond the magnitude domain
END_IF
IF ABS(fMaxBiasPct) > DL_GB_MAG_MAX THEN
    _bBadIn := TRUE;                               // 偏置上限超幅值域 | bias limit beyond the magnitude domain
END_IF
IF ABS(fDerateRatio) > DL_GB_MAG_MAX THEN
    _bBadIn := TRUE;                               // 降额倍数超幅值域 | derate multiple beyond the magnitude domain
END_IF
IF ABS(fBiasStepPct) > DL_GB_MAG_MAX THEN
    _bBadIn := TRUE;                               // 步长超幅值域 | bias step beyond the magnitude domain
END_IF

// 段 3｜组态闸：死区与偏置上限与步长须为正，降额倍数须严格大于 1（保证降额阈值高于死区）
// segment 3, configuration gate: band, bias limit and step must be positive, the derate multiple must exceed one
IF fBalanceTolPct <= DL_GB_EPS THEN
    _bCfgBad := TRUE;                              // 死区非正：失衡判据无意义 | non-positive dead band
END_IF
IF fMaxBiasPct <= DL_GB_EPS THEN
    _bCfgBad := TRUE;                              // 偏置上限非正：钳位界非法 | non-positive bias limit
END_IF
IF fBiasStepPct <= DL_GB_EPS THEN
    _bCfgBad := TRUE;                              // 步长非正：调整永不生效 | non-positive bias step
END_IF
IF fDerateRatio <= (DL_GB_RATIO_MIN + DL_GB_EPS) THEN
    _bCfgBad := TRUE;                              // 降额倍数不大于 1：降额阈值落进死区 | derate multiple not above one
END_IF
IF tBiasPeriodMs <= T#0S THEN
    _bCfgBad := TRUE;                              // 步进周期非正：TON 无意义 | non-positive step period
END_IF

// 段 4｜失衡度与阈值（每拍全量重算，无跨拍状态驻留）
// segment 4, imbalance and thresholds, fully recomputed every scan with no cross-scan state
IF (NOT _bBadIn) AND (NOT _bCfgBad) THEN
    _fImb := ABS(fTorqueMasterPct - fTorqueSlavePct); // 失衡度 [%] = |[%] − [%]| | imbalance [%]
    _fThDerate := fBalanceTolPct * fDerateRatio;   // 降额阈值 [%] = [%] × [-] | derate threshold [%]
    _fThRecover := _fThDerate - DL_GB_HYS_PCT;     // 降额恢复阈值 [%] = [%] − [%] | derate release threshold [%]
    IF _fImb <= fBalanceTolPct THEN
        bBalanced := TRUE;                         // 失衡在死区内：判定均衡 | balanced inside the dead band
    END_IF
ELSE
    _fImb := 0.0;                                  // 闸门未过：失衡度置 0，绝不让 NaN 外泄到输出 | gated, never leak NaN downstream
    _fThDerate := 0.0;                             // 闸门未过：降额阈值置 0 [%] | derate threshold zeroed
    _fThRecover := 0.0;                            // 闸门未过：恢复阈值置 0 [%] | release threshold zeroed
END_IF

// 段 5｜定时器与沿实例无条件周期刷新（R7）；步进周期 TON 自复位（R188）
// segment 5, timers and edge instances refreshed unconditionally; the step timer is self-resetting
rtReset(CLK := bReset);
tonBias(IN := (NOT tonBias.Q) AND bEnable AND (NOT _bFaultLatch) AND (_fImb > fBalanceTolPct), PT := tBiasPeriodMs);
IF rtReset.Q THEN
    _bResetLatch := TRUE;                          // 复位沿存锁存量，段 8 统一消费 | store the reset edge, consumed in segment 8
END_IF

// 段 6｜复位沿与故障锁存（复位先执行，保证本拍新故障不被抹除，R275）
// segment 6, reset edge and fault latches; reset runs first so a same-scan fault survives
IF _bResetLatch THEN
    _bFaultLatch := FALSE;                         // 清故障锁存 | clear the fault latch
    _bBadIn := FALSE;                              // 清数据非有限成因位 | clear the non-finite cause
    _bCfgBad := FALSE;                             // 清组态非法成因位（下一拍按新参数重判）| clear the configuration cause
    _fBias := 0.0;                                 // 偏置清 0 [%]：偏置不得跨复位继承 | bias cleared, never inherited across a reset
    _eState := E_DL_BalanceState.eIdle;            // 迁相回空闲 | return to idle
END_IF
IF _bBadIn AND (NOT _bFaultLatch) THEN
    _bFaultLatch := TRUE;                          // 锁存数据非有限（独立成因）| latch the non-finite cause
    _eState := E_DL_BalanceState.eFault;           // 与锁存同拍迁相（R258）| migrate in the same scan
END_IF
IF _bCfgBad AND (NOT _bFaultLatch) THEN
    _bFaultLatch := TRUE;                          // 锁存组态非法（独立成因）| latch the configuration cause
    _eState := E_DL_BalanceState.eFault;           // 与锁存同拍迁相（R258）| migrate in the same scan
END_IF

// 段 7｜主状态机：ENUM + CASE + ELSE 兜底（R6）；偏置步进只在 eBiasAdj 相内执行
// segment 7, main state machine with ENUM + CASE + ELSE fallback; bias stepping runs only inside eBiasAdj
CASE _eState OF
E_DL_BalanceState.eIdle:
    fSpeedScalePct := 0.0;                         // 空闲相速度比例 0 [%] | idle phase keeps the scale at zero
    _fBias := 0.0;                                 // 空闲相偏置清 0 [%]：不带偏置待机 | idle phase holds no bias
    // 拍 N 进入：首扫、复位沿或失能；本拍行为：偏置与放行均清 0，拒绝步进；
    // 拍 N+1 转出：使能且组态合法且数据有限 → eBalance
    // entered on the first scan, the reset edge or on disable; both the bias and the release are zeroed;
    // exits to eBalance once enabled with legal configuration and finite data
    IF bEnable AND (NOT _bCfgBad) AND (NOT _bBadIn) AND (NOT _bFaultLatch) THEN
        _eState := E_DL_BalanceState.eBalance;
    END_IF

E_DL_BalanceState.eBalance:
    fSpeedScalePct := DL_GB_SCALE_FULL;            // 均衡相满速 100 [%] | balanced phase runs at full scale
    IF NOT bEnable THEN
        _eState := E_DL_BalanceState.eIdle;         // 失能回空闲（偏置随之清 0）| disable returns to idle and clears the bias
    ELSIF _fImb > _fThDerate THEN
        _eState := E_DL_BalanceState.eDerate;       // 恶化到降额带 | worsen into the derate band
    ELSIF _fImb > fBalanceTolPct THEN
        _eState := E_DL_BalanceState.eBiasAdj;      // 超出死区：进偏置调整相 | outside the dead band, adjust the bias
    END_IF

E_DL_BalanceState.eBiasAdj:
    fSpeedScalePct := DL_GB_SCALE_FULL;            // 调整相仍满速 100 [%] | the adjustment phase still runs at full scale
    IF NOT bEnable THEN
        _eState := E_DL_BalanceState.eIdle;         // 失能回空闲 | disable returns to idle
    ELSIF _fImb > _fThDerate THEN
        _eState := E_DL_BalanceState.eDerate;       // 恶化到降额带（本相不再步进）| worsen into the derate band, stepping stops
    ELSIF _fImb <= fBalanceTolPct THEN
        _eState := E_DL_BalanceState.eBalance;      // 回到死区内：停步进，偏置保持 | back inside the band, bias held
    ELSE
        IF tonBias.Q THEN
            // 死区内不动作：此分支只在 _fImb > fBalanceTolPct 时可达，死区由上层判据与 TON 的 IN 双重保证
            // no action inside the dead band: this branch is reachable only above the band, guarded twice
            IF fTorqueMasterPct > fTorqueSlavePct THEN
                _fBias := _fBias + fBiasStepPct;    // 主轴出力偏大 → 增加从动侧偏置 [%] | master carries more, raise the slave bias
            ELSE
                _fBias := _fBias - fBiasStepPct;    // 从动侧出力偏大 → 减小偏置 [%] | slave carries more, lower the bias
            END_IF
            _fBias := ClampBias(_fBias, fMaxBiasPct); // 钳位在 ±fMaxBiasPct [%] | clamp the bias [%]
        END_IF
    END_IF

E_DL_BalanceState.eDerate:
    // 降额比例：失衡从降额阈值升到 2 倍降额阈值的过程中，速度比例从 100 线性降到 50 并饱和
    // derate scale: linear descent from 100 to 50 while the imbalance runs from the threshold to twice the threshold
    _fDen := _fThDerate;                           // 归一除子 [%] | normalisation divisor [%]
    IF _fDen > DL_GB_EPS THEN
        _fRto := (_fImb - _fThDerate) / _fDen;      // 归一比例 [-] = [%] ÷ [%]，先判零再除 | guarded division
    ELSE
        _fRto := 1.0;                              // 除子退化（组态闸已禁）→ 保守取饱和比例 | degenerate divisor, take saturation
    END_IF
    _fRto := ClampBias(_fRto, DL_GB_RATIO_MIN);    // 归一比例先钳到 [−1,1]（限值取 1.0）| clamp the ratio into the unit band
    IF _fRto < 0.0 THEN
        _fRto := 0.0;                              // 下限再钳：滞回带内不得反向抬高速度比例 | lower clamp, never raise the scale
    END_IF
    fSpeedScalePct := DL_GB_SCALE_FULL - (DL_GB_SCALE_FULL - DL_GB_SCALE_MIN) * _fRto; // [%] − [%] × [-] | derated scale [%]
    IF NOT bEnable THEN
        _eState := E_DL_BalanceState.eIdle;         // 失能回空闲 | disable returns to idle
    ELSIF _fImb <= _fThRecover THEN
        IF _fImb <= fBalanceTolPct THEN
            _eState := E_DL_BalanceState.eBalance;  // 已回到死区内 | back inside the dead band
        ELSE
            _eState := E_DL_BalanceState.eBiasAdj;  // 回到滞回带内但仍在死区外：继续调偏置 | resume bias adjustment
        END_IF
    END_IF

E_DL_BalanceState.eFault:
    fSpeedScalePct := 0.0;                         // 故障相速度比例 0 [%]，撤放行 | fault phase withdraws the release
    _fBias := 0.0;                                 // 故障相偏置清 0 [%]：安全默认不带偏置 | fault phase holds no bias
    // 驻留语义：本相只能由段 6 的复位沿迁出（唯一解除路径）；成因经 _bBadIn / _bCfgBad 分别观测
    // dwell semantics: left only through the reset edge in segment 6; causes observed via _bBadIn and _bCfgBad

ELSE
    // 非法枚举值（越界或未定义成员）：不猜，清偏置与放行并回故障相
    // illegal enumerator: no guessing, clear the bias and the release, then return to the fault phase
    fSpeedScalePct := 0.0;
    _fBias := 0.0;
    _bFaultLatch := TRUE;
    _eState := E_DL_BalanceState.eFault;
END_CASE;

// 段 8｜出口单点映射（偏置与放行在本段统一对外，CASE 后不再无条件清零 CASE 内写入量，R187）
// segment 8, single-point output mapping; nothing written inside the CASE is cleared afterwards
eState := _eState;                                 // 状态映射 | state mapping
fImbalancePct := _fImb;                            // 失衡度映射 [%] | imbalance mapping [%]
fBiasOutPct := _fBias;                             // 偏置映射 [%] | bias mapping [%]
bFaultOut := _bFaultLatch;                         // 故障锁存回放 | replay the fault latch
bCfgErr := _bCfgBad;                               // 组态非法诊断位 | bad-configuration diagnostic
bDataErr := _bBadIn;                               // 数据非有限诊断位 | non-finite data diagnostic
IF _bFaultLatch THEN
    fBiasOutPct := 0.0;                            // 故障锁存期间偏置强制 0 [%]（安全默认双保险）| bias forced to zero while latched
END_IF

// 段 9｜本拍消费量收尾（仅清沿锁存；不触碰任何锁存位与 CASE 内写入量）
// segment 9, end-of-scan cleanup; only the edge latch is cleared
_bResetLatch := FALSE;
END_FUNCTION_BLOCK

(* ---- FB_DL_GantrySkewMonitor.st ---- *)
(*==============================================================================
 * 组件名称 (Component)  : FB_DL_GantrySkewMonitor
 * 所属子库 (Sublibrary) : DL_Motion
 * 当前版本 (Version)    : 1.0.0
 * 兼容性   (Platform)   : CODESYS 3.5+ / TwinCAT 3 / 汇川 InoProShop / 施耐德 Machine Expert
 *                         仅依赖 Standard.library（TON / R_TRIG / ABS / ATAN），零厂商私有库
 * 功能描述 (Function)   : 龙门双侧偏斜监控，位置差量与角度双出口、超限分预警/报警两档。
 *                           ① 位置差量 fSkewPos = fPosLeft − fPosRight（带符号，右驱超前者为负）；
 *                           ② 角度 fSkewDeg = ATAN(fSkewPos / fGantryWidth) × 180 / π（度，带符号）。
 *                              单参 ATAN 而非 ATAN2：fGantryWidth 已过正数硬闸（> DL_GSK_EPS），
 *                              且工程上 |偏斜| 远小于 90°，该域内 ATAN(y/x) 与 ATAN2(y,x) 等价；
 *                              避开 ATAN2 在各平台库中可用性不一致的问题（跨平台可移植要求）。
 *                           ③ 双档：位置差或角度任一越预警线 → 维护级预警（bWarn，当拍量）；
 *                              任一越报警线且持续 tConfirm → 故障锁存（bAlarm，锁存至复位）。
 *                              两档并列判，取"或"关系，因为机械上位置超限与角度超限是同一次
 *                              扭曲的两种量纲表达，任一口径报警都必须报（宁可双报，不可漏报）。
 * 接口     (Interface)  : 输入 fPosLeft / fPosRight 两侧位置、fGantryWidth 两驱间距（mm，> 0）、
 *                         fSkewWarnPos / fSkewAlarmPos 位置档阈值（mm，> 0）、fSkewWarnDeg /
 *                         fSkewAlarmDeg 角度档阈值（度，> 0）、tConfirm 报警确认时间、bReset 复位；
 *                         输出 fSkewPos 差量、fSkewDeg 角度、bWarn 预警、bAlarm 报警锁存、
 *                         eState / eCause / bError。
 * 边界     (Boundary)   : ① 组态闸（覆盖每个参与判据的引脚，缺一即该判据静默失效）：
 *                         fGantryWidth <= DL_GSK_EPS（防除零把角度算成 ±Inf 或 NaN）、
 *                         位置与角度阈值 <= 0.0、报警阈值 <= 预警阈值、tConfirm <= T#0S、
 *                         任一浮点引脚 NaN（NaN 会让 ABS 比较恒假，双档同时静默失效）→ 故障锁存。
 *                         ② **本件不输出纠偏量、不发补偿指令**：龙门纠偏（如双驱转矩分配、
 *                         从动侧位置补偿）属运动学层，本件只出诊断结论。
 *                         ③ 角度换算用常量 DL_GSK_RAD2DEG，不由调用方传入（避免与本件阈值口径漂移）。
 *                         ④ TON 一枚 + R_TRIG 一枚段 0 无条件周期刷新。
 *                         ⑤ 故障相迁出唯一路径 = bReset 上升沿（R228B）。
 *                         ⑥ 零全局耦合（无 GVL / 无 VAR_EXTERNAL / 无物理地址）。
 * 分工声明 (Scope)      : 与 `FB_DL_GantrySyncAxis`（双轴同步偏差与同步控制）分工——那件关心
 *                         "同步得上不上"，可能含补偿；本件只做**偏斜监控与分档告警**，纯诊断件。
 * 来源标签 (Source Tag) : T1-6 ◐（开源参考：龙门偏斜双口径监控阈值参数域，零代码行复制）
 * 解除式   (Release)    : bReset 上升沿 ∧ 组态合法 ∧ 当拍 |fSkewPos| <= fSkewWarnPos ∧
 *                         当拍 |fSkewDeg| <= fSkewWarnDeg（回落到预警带内，R240 全当拍量）。
 *                         自证可满足：四个因子均为当拍量，龙门回到对正位置即满足，无死锁。
 * 码表     (Codes)      : 本件不占用任何全局数字码位。出口为 BOOL（bWarn / bAlarm / bError）+
 *                         ENUM（eLevel 可另读 eState / eCause）；数字码位待主控收口阶段统一派号。
 * 红线自检 (Redline)    : R1 ✓ 零 GVL/VAR_EXTERNAL ｜ R2 ✓ 零 %I/%Q/%M ｜ R3 ✓ 纯 IEC 61131-3
 *                         R4 ✓ 除零闸 + 阈值几何闸 + 浮点容差比较 ｜ R5 ✓ 声明逐行同行双语注释
 *                         R6 ✓ ENUM+CASE 含 ELSE ｜ R7 ✓ TON/R_TRIG 段 0 无条件刷新
 * 修订历史 (Revision)   : 2026-11-19  v1.0.0  R46 首版（批次 2 · 序号 7）
 *==============================================================================*)

TYPE E_DL_GskState :
(
    eIdle  := 0,    // 首拍未取到可信输入 / Awaiting trustworthy input
    eRun   := 10,   // 偏斜监控运行相 / Skew monitoring phase
    eFault := 90    // 报警锁存相（仅复位沿可迁出） / Alarm latched phase
);
END_TYPE

TYPE E_DL_GskCause :
(
    eNone       := 0,   // 无异常 / No anomaly
    eCfgIllegal := 1,   // 组态非法（宽度非正/阈值倒置/非有限） / Illegal configuration
    ePosLimit   := 2,   // 位置差量越报警线且确认窗到 / Position skew over limit confirmed
    eAngLimit   := 3,   // 角度越报警线且确认窗到 / Angle skew over limit confirmed
    ePhaseBad   := 4    // 非法相位兜底 / Illegal phase fallback
);
END_TYPE

FUNCTION_BLOCK FB_DL_GantrySkewMonitor
VAR_INPUT
    fPosLeft     : REAL := 0.0;      // 左侧（主动侧）位置 [mm] / Left, master-side position [mm]
    fPosRight    : REAL := 0.0;      // 右侧（从动侧）位置 [mm] / Right, follower-side position [mm]
    fGantryWidth : REAL := 1000.0;   // 两驱间距，域 > DL_GSK_EPS（角度换算分母） [mm] / Drive spacing, angle denominator, > epsilon [mm]
    fSkewWarnPos : REAL := 0.5;      // 位置差预警线，域 > 0.0 [mm] / Position skew warning line, > 0.0 [mm]
    fSkewAlarmPos: REAL := 2.0;      // 位置差报警线，域 > fSkewWarnPos [mm] / Position skew alarm line, > warning [mm]
    fSkewWarnDeg : REAL := 0.05;     // 角度预警线，域 > 0.0 [度] / Angle warning line, > 0.0 [deg]
    fSkewAlarmDeg: REAL := 0.20;     // 角度报警线，域 > fSkewWarnDeg [度] / Angle alarm line, > warning [deg]
    tConfirm     : TIME := T#200MS;  // 报警确认时间，域 > T#0S [ms] / Alarm confirm time, > T#0S [ms]
    bReset       : BOOL := FALSE;    // 复位，上升沿清报警锁存 [-] / Reset, rising edge clears the alarm latch
END_VAR
VAR_OUTPUT
    fSkewPos : REAL;                // 位置差量（左 − 右，带符号） [mm] / Position skew, left minus right [mm]
    fSkewDeg : REAL;                // 偏斜角度（带符号，右驱超前为负） [度] / Skew angle in degrees [deg]
    bWarn    : BOOL;                // 维护级预警（未达报警） [-] / Maintenance warning below alarm level
    bAlarm   : BOOL;                // 报警锁存 [-] / Latched alarm
    eState   : E_DL_GskState;       // 状态出口 [-] / State outlet
    eCause   : E_DL_GskCause;       // 成因出口（R190 归因唯一） [-] / Cause outlet
    bError   : BOOL;                // 故障标志（报警或组态非法） [-] / Error flag
END_VAR
VAR
    _eState  : E_DL_GskState := E_DL_GskState.eIdle;    // 内部相位（CASE 唯一写入目标） / Internal phase
    _eCause  : E_DL_GskCause := E_DL_GskCause.eNone;    // 成因锁存量 / Latched cause
    tonAlarm : TON;             // 报警确认计时，段 0 无条件调用 / Alarm confirm timer
    rtReset  : R_TRIG;          // 复位沿实例，段 0 无条件调用 / Reset edge instance
    _bFault  : BOOL;            // 报警锁存位（锁存量） / Latched alarm bit
    _bCfgBad : BOOL;            // 组态非法当拍量 [-] / Illegal configuration this scan
    _bNonFin : BOOL;            // 输入非有限当拍量 [-] / Non-finite input this scan
    _bPosOver: BOOL;            // 位置差越报警线当拍量 [-] / Position skew over the alarm line
    _bAngOver: BOOL;            // 角度越报警线当拍量 [-] / Angle skew over the alarm line
    _bWarnRaw: BOOL;            // 预警判据当拍量 [-] / Raw warning criterion
    _fSkewPos: REAL;            // 当拍差量中间量 [mm] / Skew intermediate [mm]
    _fSkewDeg: REAL;            // 当拍角度中间量 [度] / Angle intermediate [deg]
END_VAR
VAR CONSTANT
    DL_GSK_EPS     : REAL := 1.0E-6;         // 浮点判零容差（宽度与阈值统一口径） [无量纲] / Float epsilon for gates
    DL_GSK_RAD2DEG : REAL := 57.2957795;     // 弧度转度常量（180/π，7 位有效） [度/弧度] / Radians to degrees constant
END_VAR

(* —— 段 0：当拍量派生（角度先算，判据后算，顺序即依赖序） —— *)
_bNonFin := (fPosLeft <> fPosLeft) OR (fPosRight <> fPosRight)          // 位置 NaN 自反判（判等禁令唯一例外） / Position NaN tests
         OR (fGantryWidth <> fGantryWidth) OR (fSkewWarnPos <> fSkewWarnPos)
         OR (fSkewAlarmPos <> fSkewAlarmPos) OR (fSkewWarnDeg <> fSkewWarnDeg)
         OR (fSkewAlarmDeg <> fSkewAlarmDeg);                            // 阈值引脚 NaN 全量判 / Threshold NaN tests, all pins
_bCfgBad := (ABS(fGantryWidth) <= DL_GSK_EPS)                           // 宽度除零闸（缺此即角度判据静默失效） / Width divide gate
         OR (fSkewWarnPos <= 0.0) OR (fSkewAlarmPos <= fSkewWarnPos)     // 位置档几何闸 / Position threshold geometry
         OR (fSkewWarnDeg <= 0.0) OR (fSkewAlarmDeg <= fSkewWarnDeg)     // 角度档几何闸 / Angle threshold geometry
         OR (tConfirm <= T#0S) OR _bNonFin;                              // 时间闸 + 非有限 / Time gate and non-finite
_fSkewPos := fPosLeft - fPosRight;                                      // 位置差量（左 − 右） / Position skew, left minus right
IF ABS(fGantryWidth) > DL_GSK_EPS THEN                                  // 除零闸（双保险：段 0 已闸，此处防类型级直除） / Divide guard, second layer
    _fSkewDeg := ATAN(_fSkewPos / fGantryWidth) * DL_GSK_RAD2DEG;       // 角度换算：单参 ATAN，宽度为正故符号随差量 / Angle via single-arg ATAN, sign follows skew
ELSE
    _fSkewDeg := 0.0;                                                   // 宽度病态：角度不宣称 / Degenerate width: angle not claimed
END_IF
_bPosOver := ABS(_fSkewPos) > fSkewAlarmPos;                            // 位置差越报警线 / Position skew over the alarm line
_bAngOver := ABS(_fSkewDeg) > fSkewAlarmDeg;                            // 角度越报警线 / Angle skew over the alarm line
_bWarnRaw := (ABS(_fSkewPos) > fSkewWarnPos) OR (ABS(_fSkewDeg) > fSkewWarnDeg);   // 预警判据（双口径取或） / Warning criterion, either unit
rtReset(CLK := bReset);                                                 // 复位沿，每拍必调（R228A） / Reset edge, every scan
tonAlarm(IN := _bPosOver OR _bAngOver, PT := tConfirm);                 // 报警确认窗（IN 由当拍判据派生） / Alarm confirm window

(* —— 段 1：单拍量预清零（锁存量 _bFault / _eCause 不入清单，R107） —— *)
fSkewPos := 0.0;        // 差量出口每拍预清，段 6 回填 / Skew outlet preset
fSkewDeg := 0.0;        // 角度出口每拍预清 / Angle outlet preset
bWarn    := FALSE;      // 预警位每拍预清 / Warning preset
bAlarm   := FALSE;      // 报警出口每拍预清，锁存分支同拍回填 / Alarm outlet preset
bError   := FALSE;      // 故障标志每拍预清（R45 配对） / Error flag preset

(* —— 段 2：复位沿 + 组态闸 —— *)
IF rtReset.Q THEN
    _bFault := FALSE;                                   // 清报警锁存（锁存量） / Clear the alarm latch
    _eCause := E_DL_GskCause.eNone;                      // 清成因 / Clear cause
    IF _eState = E_DL_GskState.eFault THEN
        _eState := E_DL_GskState.eIdle;                  // 故障相迁出（R228B） / Leave fault phase
    END_IF
END_IF
IF _bCfgBad THEN
    _bFault := TRUE;                                     // 组态非法锁存 / Latch illegal configuration
    _eCause := E_DL_GskCause.eCfgIllegal;                // 归因：组态非法 / Cause: illegal configuration
    bError  := TRUE;                                     // 故障标志同拍置位 / Error flag set same scan
END_IF

(* —— 段 3：报警分级（位置与角度归因分开，先位置后角度，同拍双越限时归因确定） —— *)
IF (NOT _bFault) AND (NOT _bCfgBad) AND tonAlarm.Q THEN
    _bFault := TRUE;                                     // 锁存 / Latch
    IF _bPosOver THEN
        _eCause := E_DL_GskCause.ePosLimit;              // 归因：位置差越限（优先） / Cause: position skew over limit
    ELSE
        _eCause := E_DL_GskCause.eAngLimit;              // 归因：角度越限 / Cause: angle skew over limit
    END_IF
    bError := TRUE;                                      // 故障标志同拍置位 / Error flag set same scan
END_IF

(* —— 段 4：预警（维护级，不锁存；报警命中时不再宣称预警） —— *)
IF (NOT _bFault) AND _bWarnRaw THEN
    bWarn := TRUE;                                       // 维护级预警 / Maintenance warning
END_IF

(* —— 段 5：锁存相位迁移闸 —— *)
IF _bFault AND (_eState <> E_DL_GskState.eFault) THEN
    _eState := E_DL_GskState.eFault;                     // 锁存即入故障相 / Latch enters fault phase
END_IF

(* —— 段 6：相位机（ENUM 全成员显式标签 + ELSE 兜底，R128） —— *)
CASE _eState OF

E_DL_GskState.eIdle:
    IF (NOT _bNonFin) AND (NOT _bCfgBad) THEN            // 出口 1：输入可信 / Input trustworthy
        _eState := E_DL_GskState.eRun;
    ELSIF _bFault THEN                                   // 出口 2：故障锁存 / Fault latched
        _eState := E_DL_GskState.eFault;
    END_IF

E_DL_GskState.eRun:
    IF _bFault THEN                                      // 出口 1：报警锁存 / Alarm latched
        _eState := E_DL_GskState.eFault;
    ELSIF rtReset.Q THEN                                 // 出口 2：复位沿回观测相 / Reset edge back to observation
        _eState := E_DL_GskState.eIdle;
    END_IF

E_DL_GskState.eFault:
    ;                                                    // 故障相：仅段 2 复位沿可迁出 / Only the reset edge leaves this phase

ELSE
    _bFault := TRUE;                                     // 非法相位兜底锁存 / Illegal-phase fallback latch
    _eCause := E_DL_GskCause.ePhaseBad;                  // 归因：非法相位 / Cause: illegal phase
    _eState := E_DL_GskState.eFault;                     // 强拉故障相 / Force fault phase

END_CASE

(* —— 段 7：出口单点映射（差量与角度始终回放当拍计算值，故障相亦然——诊断量不可清零） —— *)
fSkewPos := _fSkewPos;                                   // 差量出口 / Skew outlet
fSkewDeg := _fSkewDeg;                                   // 角度出口 / Angle outlet
bAlarm   := _bFault;                                     // 报警与锁存同源（R191） / Alarm from latch
bError   := _bFault OR _bCfgBad;                         // 故障标志 = 锁存或组态非法 / Error = latch or illegal config
IF _bFault THEN
    bWarn := FALSE;                                      // 报警相不再宣称「仅预警」 / No warning claim in alarm
END_IF
eState := _eState;                                       // 状态出口 / State outlet
eCause := _eCause;                                       // 成因出口 / Cause outlet

END_FUNCTION_BLOCK
